(* IEC 61131-3 sources: canworks/library/modbus, 29 files *)

(* ---- CW_CHAR.st ---- *)
FUNCTION CW_CHAR : STRING
(* The one-character STRING of byte CODE ('' for 0), for building a STRING
   from bytes in plain ST: a look-up in tables of every byte value, 32 per
   table so that each fits the shortest default STRING length. *)
VAR_INPUT
  CODE : BYTE;
END_VAR
VAR
  t0 : STRING := '$01$02$03$04$05$06$07$08$09$0A$0B$0C$0D$0E$0F$10$11$12$13$14$15$16$17$18$19$1A$1B$1C$1D$1E$1F';
  t1 : STRING := '$20$21$22$23$24$25$26$27$28$29$2A$2B$2C$2D$2E$2F$30$31$32$33$34$35$36$37$38$39$3A$3B$3C$3D$3E$3F';
  t2 : STRING := '$40$41$42$43$44$45$46$47$48$49$4A$4B$4C$4D$4E$4F$50$51$52$53$54$55$56$57$58$59$5A$5B$5C$5D$5E$5F';
  t3 : STRING := '$60$61$62$63$64$65$66$67$68$69$6A$6B$6C$6D$6E$6F$70$71$72$73$74$75$76$77$78$79$7A$7B$7C$7D$7E$7F';
  t4 : STRING := '$80$81$82$83$84$85$86$87$88$89$8A$8B$8C$8D$8E$8F$90$91$92$93$94$95$96$97$98$99$9A$9B$9C$9D$9E$9F';
  t5 : STRING := '$A0$A1$A2$A3$A4$A5$A6$A7$A8$A9$AA$AB$AC$AD$AE$AF$B0$B1$B2$B3$B4$B5$B6$B7$B8$B9$BA$BB$BC$BD$BE$BF';
  t6 : STRING := '$C0$C1$C2$C3$C4$C5$C6$C7$C8$C9$CA$CB$CC$CD$CE$CF$D0$D1$D2$D3$D4$D5$D6$D7$D8$D9$DA$DB$DC$DD$DE$DF';
  t7 : STRING := '$E0$E1$E2$E3$E4$E5$E6$E7$E8$E9$EA$EB$EC$ED$EE$EF$F0$F1$F2$F3$F4$F5$F6$F7$F8$F9$FA$FB$FC$FD$FE$FF';
  k : INT;
END_VAR
k := BYTE_TO_INT(CODE);
CASE k / 32 OF
  0:
    IF k > 0 THEN
      CW_CHAR := MID(t0, 1, k);
    ELSE
      CW_CHAR := '';
    END_IF;
  1: CW_CHAR := MID(t1, 1, k MOD 32 + 1);
  2: CW_CHAR := MID(t2, 1, k MOD 32 + 1);
  3: CW_CHAR := MID(t3, 1, k MOD 32 + 1);
  4: CW_CHAR := MID(t4, 1, k MOD 32 + 1);
  5: CW_CHAR := MID(t5, 1, k MOD 32 + 1);
  6: CW_CHAR := MID(t6, 1, k MOD 32 + 1);
ELSE
  CW_CHAR := MID(t7, 1, k MOD 32 + 1);
END_CASE;
END_FUNCTION

FUNCTION CW_CHAR_CODE : BYTE
(* The byte value of the first character of C (0 for ''). *)
VAR_INPUT
  C : STRING;
END_VAR
VAR
  t0 : STRING := '$01$02$03$04$05$06$07$08$09$0A$0B$0C$0D$0E$0F$10$11$12$13$14$15$16$17$18$19$1A$1B$1C$1D$1E$1F';
  t1 : STRING := '$20$21$22$23$24$25$26$27$28$29$2A$2B$2C$2D$2E$2F$30$31$32$33$34$35$36$37$38$39$3A$3B$3C$3D$3E$3F';
  t2 : STRING := '$40$41$42$43$44$45$46$47$48$49$4A$4B$4C$4D$4E$4F$50$51$52$53$54$55$56$57$58$59$5A$5B$5C$5D$5E$5F';
  t3 : STRING := '$60$61$62$63$64$65$66$67$68$69$6A$6B$6C$6D$6E$6F$70$71$72$73$74$75$76$77$78$79$7A$7B$7C$7D$7E$7F';
  t4 : STRING := '$80$81$82$83$84$85$86$87$88$89$8A$8B$8C$8D$8E$8F$90$91$92$93$94$95$96$97$98$99$9A$9B$9C$9D$9E$9F';
  t5 : STRING := '$A0$A1$A2$A3$A4$A5$A6$A7$A8$A9$AA$AB$AC$AD$AE$AF$B0$B1$B2$B3$B4$B5$B6$B7$B8$B9$BA$BB$BC$BD$BE$BF';
  t6 : STRING := '$C0$C1$C2$C3$C4$C5$C6$C7$C8$C9$CA$CB$CC$CD$CE$CF$D0$D1$D2$D3$D4$D5$D6$D7$D8$D9$DA$DB$DC$DD$DE$DF';
  t7 : STRING := '$E0$E1$E2$E3$E4$E5$E6$E7$E8$E9$EA$EB$EC$ED$EE$EF$F0$F1$F2$F3$F4$F5$F6$F7$F8$F9$FA$FB$FC$FD$FE$FF';
  first : STRING;
  p : INT;
END_VAR
CW_CHAR_CODE := BYTE#0;
IF LEN(C) = 0 THEN
  RETURN;
END_IF;
first := LEFT(C, 1);
p := FIND(t0, first);
IF p > 0 THEN
  CW_CHAR_CODE := INT_TO_BYTE(p);
  RETURN;
END_IF;
p := FIND(t1, first);
IF p > 0 THEN
  CW_CHAR_CODE := INT_TO_BYTE(31 + p);
  RETURN;
END_IF;
p := FIND(t2, first);
IF p > 0 THEN
  CW_CHAR_CODE := INT_TO_BYTE(63 + p);
  RETURN;
END_IF;
p := FIND(t3, first);
IF p > 0 THEN
  CW_CHAR_CODE := INT_TO_BYTE(95 + p);
  RETURN;
END_IF;
p := FIND(t4, first);
IF p > 0 THEN
  CW_CHAR_CODE := INT_TO_BYTE(127 + p);
  RETURN;
END_IF;
p := FIND(t5, first);
IF p > 0 THEN
  CW_CHAR_CODE := INT_TO_BYTE(159 + p);
  RETURN;
END_IF;
p := FIND(t6, first);
IF p > 0 THEN
  CW_CHAR_CODE := INT_TO_BYTE(191 + p);
  RETURN;
END_IF;
p := FIND(t7, first);
IF p > 0 THEN
  CW_CHAR_CODE := INT_TO_BYTE(223 + p);
END_IF;
END_FUNCTION

(* ---- CW_REAL.st ---- *)
FUNCTION CW_DWORD_TO_REAL : REAL
(* The REAL whose IEEE 754 bit pattern is IN (a 32-bit value read from two
   Modbus registers). Infinities come back as +/-3.4E38, NaN as 0.0. *)
VAR_INPUT
  IN : DWORD;
END_VAR
VAR
  e : INT;
  m : LREAL;
  x : LREAL;
END_VAR
e := DWORD_TO_INT(SHR(IN, 23) AND DWORD#16#FF);
m := UDINT_TO_LREAL(DWORD_TO_UDINT(IN AND DWORD#16#7FFFFF));
IF e = 255 THEN
  IF m <> 0.0 THEN
    x := 0.0;
  ELSE
    x := 3.4028234663852886E38;
  END_IF;
ELSIF e = 0 THEN
  x := m * EXPT(2.0, -149);
ELSE
  x := (m + 8388608.0) * EXPT(2.0, e - 150);
END_IF;
IF (IN AND DWORD#16#80000000) <> DWORD#0 THEN
  x := -x;
END_IF;
CW_DWORD_TO_REAL := LREAL_TO_REAL(x);
END_FUNCTION

FUNCTION CW_REAL_TO_DWORD : DWORD
(* The IEEE 754 bit pattern of IN, to send a REAL in two Modbus registers. *)
VAR_INPUT
  IN : REAL;
END_VAR
VAR
  a : LREAL;
  e : INT;
  sign : DWORD;
END_VAR
a := REAL_TO_LREAL(IN);
sign := DWORD#0;
IF a < 0.0 THEN
  sign := DWORD#16#80000000;
  a := -a;
END_IF;
IF a <> a THEN
  CW_REAL_TO_DWORD := DWORD#16#7FC00000;
  RETURN;
END_IF;
IF a = 0.0 THEN
  CW_REAL_TO_DWORD := sign;
  RETURN;
END_IF;
IF a > 3.4028234663852886E38 THEN
  CW_REAL_TO_DWORD := sign OR DWORD#16#7F800000;
  RETURN;
END_IF;
e := LREAL_TO_INT(TRUNC(LN(a) / LN(2.0)));
WHILE a / EXPT(2.0, e) >= 2.0 DO
  e := e + 1;
END_WHILE;
WHILE a / EXPT(2.0, e) < 1.0 DO
  e := e - 1;
END_WHILE;
IF e < -126 THEN
  CW_REAL_TO_DWORD := sign OR UDINT_TO_DWORD(LREAL_TO_UDINT(a * EXPT(2.0, 149)));
ELSE
  CW_REAL_TO_DWORD := sign OR SHL(INT_TO_DWORD(e + 127), 23) OR UDINT_TO_DWORD(LREAL_TO_UDINT((a / EXPT(2.0, e) - 1.0) * 8388608.0));
END_IF;
END_FUNCTION

FUNCTION CW_LWORD_TO_LREAL : LREAL
(* The LREAL whose IEEE 754 bit pattern is IN (a 64-bit value read from four
   Modbus registers). Infinities come back as +/-1.79E308, NaN as 0.0. *)
VAR_INPUT
  IN : LWORD;
END_VAR
VAR
  e : INT;
  m : LREAL;
  x : LREAL;
END_VAR
e := LWORD_TO_INT(SHR(IN, 52) AND LWORD#16#7FF);
m := ULINT_TO_LREAL(LWORD_TO_ULINT(IN AND LWORD#16#FFFFFFFFFFFFF));
IF e = 2047 THEN
  IF m <> 0.0 THEN
    x := 0.0;
  ELSE
    x := 1.7976931348623157E308;
  END_IF;
ELSIF e = 0 THEN
  x := m * EXPT(2.0, -1074);
ELSE
  x := (m + 4503599627370496.0) * EXPT(2.0, e - 1075);
END_IF;
IF (IN AND SHL(LWORD#1, 63)) <> LWORD#0 THEN
  x := -x;
END_IF;
CW_LWORD_TO_LREAL := x;
END_FUNCTION

FUNCTION CW_LREAL_TO_LWORD : LWORD
(* The IEEE 754 bit pattern of IN, to send an LREAL in four Modbus registers. *)
VAR_INPUT
  IN : LREAL;
END_VAR
VAR
  a : LREAL;
  e : INT;
  sign : LWORD;
END_VAR
a := IN;
sign := LWORD#0;
IF a < 0.0 THEN
  sign := SHL(LWORD#1, 63);
  a := -a;
END_IF;
IF a <> a THEN
  CW_LREAL_TO_LWORD := LWORD#16#7FF8000000000000;
  RETURN;
END_IF;
IF a = 0.0 THEN
  CW_LREAL_TO_LWORD := sign;
  RETURN;
END_IF;
IF a > 1.7976931348623157E308 THEN
  CW_LREAL_TO_LWORD := sign OR LWORD#16#7FF0000000000000;
  RETURN;
END_IF;
e := LREAL_TO_INT(TRUNC(LN(a) / LN(2.0)));
WHILE a / EXPT(2.0, e) >= 2.0 DO
  e := e + 1;
END_WHILE;
WHILE a / EXPT(2.0, e) < 1.0 DO
  e := e - 1;
END_WHILE;
IF e < -1022 THEN
  CW_LREAL_TO_LWORD := sign OR ULINT_TO_LWORD(LREAL_TO_ULINT(a * EXPT(2.0, 537) * EXPT(2.0, 537)));
ELSE
  CW_LREAL_TO_LWORD := sign OR SHL(INT_TO_LWORD(e + 1023), 52) OR ULINT_TO_LWORD(LREAL_TO_ULINT((a / EXPT(2.0, e) - 1.0) * 4503599627370496.0));
END_IF;
END_FUNCTION

(* ---- CAN_BUS_INFO.st ---- *)
(*
 * CAN_BUS_INFO: the state of network NETWORK (one of the first 8) from the
 * bridge's network info block, updated every 100 ms, without a request:
 * STATE (0 error active, 1 warning, 2 error passive, 3 bus off, 4 unknown),
 * TX_ERRORS and RX_ERRORS (error counters), BUS_OFF_COUNT, BUS_LOAD (%),
 * RX_COUNT and TX_COUNT (frames), ERROR_FRAMES. ERROR_ID
 * (docs/plc-library.md#frame-blocks): 2 no such network, 20 the bridge is
 * not reachable, 22 the config has no network info (or NETWORK is past the
 * first 8).
 *)
(*
 * LINK is the generated `canworks.link` (ARRAY[0..1279] OF WORD); the block reads the bridge's network info block (see
 * CW_LINK_SERVICE for the words).
 *)
FUNCTION_BLOCK CAN_BUS_INFO
VAR_INPUT
  NETWORK : USINT;
END_VAR
VAR_IN_OUT
  LINK : ARRAY[0..1279] OF WORD;
END_VAR
VAR_OUTPUT
  STATE : USINT;
  TX_ERRORS : UINT;
  RX_ERRORS : UINT;
  BUS_OFF_COUNT : UDINT;
  BUS_LOAD : USINT;
  RX_COUNT : UDINT;
  TX_COUNT : UDINT;
  ERROR_FRAMES : UDINT;
  ERROR : BOOL;
  ERROR_ID : UINT;
END_VAR
VAR
  p : INT;
END_VAR
  ERROR_ID := 0;
  IF (LINK[21] AND WORD#16#0001) = WORD#0 THEN
    ERROR_ID := 20;
  ELSIF (LINK[89] AND WORD#16#0020) = WORD#0 OR NETWORK > 7 THEN
    ERROR_ID := 22;
  ELSE
    p := 960 + 18 * USINT_TO_INT(NETWORK);
    IF LINK[p + 17] = WORD#0 THEN
      ERROR_ID := 2;
    END_IF;
  END_IF;
  ERROR := ERROR_ID <> 0;
  IF ERROR THEN
    STATE := 4;
    TX_ERRORS := 0;
    RX_ERRORS := 0;
    BUS_OFF_COUNT := 0;
    BUS_LOAD := 0;
    RX_COUNT := 0;
    TX_COUNT := 0;
    ERROR_FRAMES := 0;
    RETURN;
  END_IF;
  STATE := WORD_TO_USINT(SHR(LINK[p], 8));
  BUS_LOAD := WORD_TO_USINT(LINK[p] AND WORD#16#00FF);
  TX_ERRORS := WORD_TO_UINT(LINK[p + 1]);
  RX_ERRORS := WORD_TO_UINT(LINK[p + 2]);
  BUS_OFF_COUNT := WORD_TO_UDINT(LINK[p + 3]) * 65536 + WORD_TO_UDINT(LINK[p + 4]);
  RX_COUNT := WORD_TO_UDINT(LINK[p + 5]) * 65536 + WORD_TO_UDINT(LINK[p + 6]);
  TX_COUNT := WORD_TO_UDINT(LINK[p + 7]) * 65536 + WORD_TO_UDINT(LINK[p + 8]);
  ERROR_FRAMES := WORD_TO_UDINT(LINK[p + 9]) * 65536 + WORD_TO_UDINT(LINK[p + 10]);
END_FUNCTION_BLOCK

(* ---- CAN_RECEIVE.st ---- *)
(*
 * CAN_RECEIVE: receives the CAN frames of network NETWORK whose identifier
 * matches ID under MASK (MASK 0: ID exactly; ALL_IDS: every frame of that
 * format), standard or EXTENDED, through a receiver of the bridge with a
 * queue of DEPTH frames (0: 32, at most 256). ENABLE opens it. Each call
 * gives at most one frame, oldest first: RECEIVED with RX_ID, RX_EXTENDED,
 * RX_RTR, RX_DLC, RX_DATA and TIMESTAMP (UTC microseconds, the receive time
 * of the bridge's batch, which its frames share: about one poll); call it
 * again in the same scan to read more
 * (`WHILE rx.RECEIVED DO ... rx(...); END_WHILE`).
 * QUEUED frames still wait in the bridge, OVERFLOW the queue was full,
 * DROPPED frames lost. ERROR_ID (docs/plc-library.md#frame-blocks): 1 the
 * network is not running, 2 no such network, 3 invalid input, 5 no free
 * receiver, 8 the bridge closed the receiver (it opens again), 20 the
 * bridge is not reachable, 22 the config has no receive or request mailbox.
 * After 1, 8 and 20 it opens again by itself.
 *)
(*
 * LINK is the generated `canworks.link` (ARRAY[0..1279] OF WORD); the block uses the bridge's receive mailbox and, to open and close its receiver, a
 * request mailbox (see
 * CW_LINK_SERVICE for the words).
 *)
FUNCTION_BLOCK CAN_RECEIVE
VAR_INPUT
  ENABLE : BOOL;
  NETWORK : USINT;
  ID : UDINT;
  MASK : UDINT;
  ALL_IDS : BOOL;
  EXTENDED : BOOL;
  DEPTH : UINT;
END_VAR
VAR_IN_OUT
  RX_DATA : ARRAY[0..7] OF BYTE;
  LINK : ARRAY[0..1279] OF WORD;
END_VAR
VAR_OUTPUT
  ACTIVE : BOOL;
  RECEIVED : BOOL;
  RX_ID : UDINT;
  RX_EXTENDED : BOOL;
  RX_RTR : BOOL;
  RX_DLC : USINT;
  TIMESTAMP : ULINT;
  QUEUED : UINT;
  OVERFLOW : BOOL;
  DROPPED : UDINT;
  ERROR : BOOL;
  ERROR_ID : UINT;
END_VAR
VAR
  rx : CW_RX;
  prev : BOOL;
  was_active : BOOL;
  last_drop : WORD;
  id_mask : UDINT;
  rec : INT;
  i : INT;
END_VAR
  IF ENABLE AND NOT prev THEN
    QUEUED := 0;
    OVERFLOW := FALSE;
    DROPPED := 0;
  END_IF;
  prev := ENABLE;
  IF ALL_IDS THEN
    id_mask := 0;
  ELSIF MASK <> 0 THEN
    id_mask := MASK;
  ELSIF EXTENDED THEN
    id_mask := 16#1FFFFFFF;
  ELSE
    id_mask := 16#7FF;
  END_IF;
  rx(ENABLE := ENABLE, CHANGED := FALSE, NEXT := TRUE, KIND := 1, NETWORK := NETWORK,
     FLAGS := SEL(EXTENDED, USINT#0, USINT#1), DEPTH := DEPTH, ID := ID, MASK := id_mask, RETRY := DWORD#16#00100102,
     LINK := LINK);
  IF rx.ACTIVE AND NOT was_active THEN
    last_drop := WORD#0;
  END_IF;
  was_active := rx.ACTIVE;
  RECEIVED := rx.RECEIVED;
  IF RECEIVED THEN
    rec := rx.REC;
    QUEUED := WORD_TO_UINT(LINK[rec + 1]);
    DROPPED := DROPPED + WORD_TO_UDINT(DINT_TO_WORD(WORD_TO_DINT(LINK[rec + 2]) - WORD_TO_DINT(last_drop)));
    last_drop := LINK[rec + 2];
    OVERFLOW := (LINK[rec] AND WORD#16#0004) <> WORD#0;
    TIMESTAMP := LWORD_TO_ULINT(SHL(WORD_TO_LWORD(LINK[741]), 48) OR SHL(WORD_TO_LWORD(LINK[742]), 32) OR
                 SHL(WORD_TO_LWORD(LINK[743]), 16) OR WORD_TO_LWORD(LINK[744]));
    RX_ID := WORD_TO_UDINT(LINK[rec + 3]) * 65536 + WORD_TO_UDINT(LINK[rec + 4]);
    RX_EXTENDED := (LINK[rec + 5] AND WORD#16#0100) <> WORD#0;
    RX_RTR := (LINK[rec + 5] AND WORD#16#0200) <> WORD#0;
    RX_DLC := WORD_TO_USINT(LINK[rec + 5] AND WORD#16#00FF);
    FOR i := 0 TO 3 DO
      RX_DATA[2 * i] := WORD_TO_BYTE(SHR(LINK[rec + 6 + i], 8));
      RX_DATA[2 * i + 1] := WORD_TO_BYTE(LINK[rec + 6 + i]);
    END_FOR;
  END_IF;
  ACTIVE := rx.ACTIVE;
  ERROR := rx.ERROR;
  ERROR_ID := rx.ERROR_ID;
END_FUNCTION_BLOCK

(* ---- CAN_SEND.st ---- *)
(*
 * CAN_SEND: sends one CAN frame (ID, EXTENDED, RTR, DLC 0..8 bytes of DATA)
 * on network NETWORK. A rising edge of EXECUTE starts it; BUSY until the
 * bridge has sent it, then DONE or ERROR with ERROR_ID
 * (docs/plc-library.md#frame-blocks): 1 the network is not running, 2 no
 * such network, 3 invalid input, 5 too many frames wait, 6 not sent within
 * TIMEOUT (T#0s: 1 s), 7 the bus is off, 8 cancelled, 20 the bridge is not
 * reachable, 22 the config has no request mailbox.
 *)
(*
 * LINK is the generated `canworks.link` (ARRAY[0..1279] OF WORD); the block uses a request mailbox of the bridge (`mailboxes` in the config); instances share
 * them in the order they started (see
 * CW_LINK_SERVICE for the words).
 *)
FUNCTION_BLOCK CAN_SEND
VAR_INPUT
  EXECUTE : BOOL;
  NETWORK : USINT;
  ID : UDINT;
  EXTENDED : BOOL;
  RTR : BOOL;
  DLC : USINT;
  TIMEOUT : TIME;
END_VAR
VAR_IN_OUT
  DATA : ARRAY[0..7] OF BYTE;
  LINK : ARRAY[0..1279] OF WORD;
END_VAR
VAR_OUTPUT
  BUSY : BOOL;
  DONE : BOOL;
  ERROR : BOOL;
  ERROR_ID : UINT;
END_VAR
VAR
  x : CW_REQUEST;
  buf : ARRAY[0..1784] OF BYTE;
  prev : BOOL;
  refused : UINT;
  flags : WORD;
  ms : UDINT;
  i : INT;
END_VAR
  IF EXECUTE AND NOT prev AND NOT x.BUSY THEN
    refused := 0;
    IF DLC > 8 THEN
      refused := 3;
    END_IF;
    FOR i := 0 TO 7 DO
      buf[i] := DATA[i];
    END_FOR;
  ELSIF NOT EXECUTE THEN
    refused := 0;
  END_IF;
  prev := EXECUTE;
  flags := SEL(EXTENDED, WORD#0, WORD#1) OR SEL(RTR, WORD#0, WORD#2);
  ms := DWORD_TO_UDINT(TIME_TO_DWORD(TIMEOUT));
  IF ms > 65535 THEN
    ms := 65535;
  END_IF;
  x(EXECUTE := EXECUTE AND refused = 0, OP := 5, NET := NETWORK, A0 := DWORD_TO_WORD(SHR(UDINT_TO_DWORD(ID), 16)),
    A1 := UDINT_TO_WORD(ID), A2 := SHL(flags, 8) OR USINT_TO_WORD(DLC), A3 := UDINT_TO_WORD(ms), A4 := WORD#0, A5 := WORD#0,
    LENGTH := 8, FETCH_MAX := 0, LINK := LINK, DATA := buf);
  BUSY := x.BUSY;
  DONE := x.DONE;
  ERROR := x.ERROR OR refused <> 0;
  ERROR_ID := SEL(refused <> 0, x.ERROR_ID, refused);
END_FUNCTION_BLOCK

(* ---- CAN_SEND_CYCLIC.st ---- *)
(*
 * CAN_SEND_CYCLIC: the bridge sends one CAN frame (ID, EXTENDED, DLC bytes
 * of DATA) on network NETWORK every PERIOD (1 ms .. 60 s) while ENABLE is
 * TRUE. Changed DATA, DLC or PERIOD go to the bridge when they change; the
 * block must be called at least every second (its keepalive), or the bridge
 * stops the frame. ACTIVE while the job runs, COUNT frames sent. ERROR_ID
 * (docs/plc-library.md#frame-blocks): 1 the network is not running, 2 no
 * such network, 3 invalid input, 5 no free cyclic job, 7 the bus is off
 * (the job stays), 8 cancelled (the bridge stopped the job; it starts
 * again), 20 the bridge is not reachable, 22 the config has no request
 * mailbox or no cyclic jobs. After 1, 7, 8 and 20 it starts again by itself.
 *)
(*
 * LINK is the generated `canworks.link` (ARRAY[0..1279] OF WORD); the block uses a request mailbox of the bridge (`mailboxes` in the config); instances share
 * them in the order they started, and a cyclic job of the bridge's table (see
 * CW_LINK_SERVICE for the words).
 *)
FUNCTION_BLOCK CAN_SEND_CYCLIC
VAR_INPUT
  ENABLE : BOOL;
  NETWORK : USINT;
  ID : UDINT;
  EXTENDED : BOOL;
  DLC : USINT;
  PERIOD : TIME;
END_VAR
VAR_IN_OUT
  DATA : ARRAY[0..7] OF BYTE;
  LINK : ARRAY[0..1279] OF WORD;
END_VAR
VAR_OUTPUT
  ACTIVE : BOOL;
  COUNT : UDINT;
  ERROR : BOOL;
  ERROR_ID : UINT;
END_VAR
VAR
  mb : CW_MB_CALL;
  prev : BOOL;
  phase : USINT;           (* 0 off, 1 starting, 2 running, 3 updating, 4 stopping *)
  job : INT;
  gen : WORD;
  tick0 : WORD;
  sent : ARRAY[0..7] OF BYTE;
  sent_dlc : USINT;
  sent_ms : UDINT;
  ms : UDINT;
  changed : BOOL;
  t : INT;
  i : INT;
  err : UINT;
  fresh : BOOL;
END_VAR
  err := 0;
  ms := DWORD_TO_UDINT(TIME_TO_DWORD(PERIOD));
  IF ms > 65535 THEN
    ms := 65535;
  END_IF;
  IF ENABLE AND NOT prev THEN
    COUNT := 0;
    ERROR := FALSE;
    ERROR_ID := 0;
  END_IF;
  IF (LINK[21] AND WORD#16#0001) = WORD#0 AND phase <> 0 THEN
    mb(RUN := FALSE, LINK := LINK);
    phase := 0;
    IF ENABLE THEN
      err := 20;
    END_IF;
  END_IF;
  IF phase = 2 OR phase = 3 THEN
    LINK[128 + job] := UDINT_TO_WORD(WORD_TO_UDINT(LINK[128 + job]) + 1);
    t := 1105 + 4 * job;
    fresh := (DINT_TO_WORD(WORD_TO_DINT(LINK[1104]) - WORD_TO_DINT(tick0)) AND WORD#16#8000) = WORD#0;
    IF fresh AND LINK[t + 1] <> gen THEN
      mb(RUN := FALSE, LINK := LINK);
      phase := 0;
      err := 8;
    ELSIF fresh THEN
      COUNT := WORD_TO_UDINT(LINK[t + 2]) * 65536 + WORD_TO_UDINT(LINK[t + 3]);
      IF SHR(LINK[t], 8) = WORD#2 THEN
        ERROR := TRUE;
        ERROR_ID := WORD_TO_UINT(LINK[t] AND WORD#16#00FF);
      ELSIF ERROR AND ERROR_ID = 7 THEN
        ERROR := FALSE;
        ERROR_ID := 0;
      END_IF;
    END_IF;
  END_IF;
  IF (phase = 2 OR phase = 3) AND NOT ENABLE THEN
    phase := 4;
  END_IF;
  changed := DLC <> sent_dlc OR ms <> sent_ms;
  FOR i := 0 TO 7 DO
    IF DATA[i] <> sent[i] THEN
      changed := TRUE;
    END_IF;
  END_FOR;
  IF phase = 2 AND changed THEN
    phase := 3;
  END_IF;
  IF phase = 0 AND ENABLE AND err = 0 AND
     NOT (ERROR AND ERROR_ID <> 1 AND ERROR_ID <> 7 AND ERROR_ID <> 8 AND ERROR_ID <> 20) THEN
    ERROR := FALSE;
    ERROR_ID := 0;
    IF (LINK[21] AND WORD#16#0001) = WORD#0 THEN
      err := 20;
    ELSIF (LINK[89] AND WORD#16#0007) = WORD#0 OR (LINK[89] AND WORD#16#1F00) = WORD#0 THEN
      err := 22;
    ELSIF DLC > 8 THEN
      err := 3;
    ELSE
      phase := 1;
    END_IF;
  END_IF;
  IF phase = 1 OR phase = 3 OR phase = 4 THEN
    mb(RUN := TRUE, SEND := FALSE, LINK := LINK);
    IF mb.LOST THEN
      phase := 0;
      err := SEL(ENABLE, UINT#0, UINT#20);
    ELSIF mb.ANSWERED THEN
      IF phase = 4 THEN
        phase := 0;
      ELSIF mb.ERR <> 0 THEN
        err := mb.ERR;
        IF phase = 1 OR mb.ERR = 8 THEN
          phase := 0;
        ELSE
          phase := 2;
        END_IF;
      ELSE
        IF phase = 1 THEN
          job := WORD_TO_INT(LINK[mb.BASE + 74]);
          gen := LINK[mb.BASE + 75];
          tick0 := LINK[mb.BASE + 76];
          COUNT := 0;
        END_IF;
        phase := 2;
      END_IF;
      mb(RUN := FALSE, LINK := LINK);
    ELSIF mb.OWNED AND NOT mb.WAITING THEN
      IF phase = 4 THEN
        mb(RUN := TRUE, SEND := TRUE, OP := 7, NET := NETWORK, A0 := INT_TO_WORD(job), A1 := WORD#0, A2 := WORD#0, A3 := WORD#0,
           A4 := WORD#0, A5 := WORD#0, LINK := LINK);
      ELSE
        FOR i := 0 TO 3 DO
          LINK[mb.BASE + 8 + i] := SHL(BYTE_TO_WORD(DATA[2 * i]), 8) OR BYTE_TO_WORD(DATA[2 * i + 1]);
          sent[2 * i] := DATA[2 * i];
          sent[2 * i + 1] := DATA[2 * i + 1];
        END_FOR;
        sent_dlc := DLC;
        sent_ms := ms;
        mb(RUN := TRUE, SEND := TRUE, OP := 6, NET := NETWORK, A0 := SEL(phase = 1, INT_TO_WORD(job), WORD#16#FFFF),
           A1 := DWORD_TO_WORD(SHR(UDINT_TO_DWORD(ID), 16)), A2 := UDINT_TO_WORD(ID),
           A3 := SHL(SEL(EXTENDED, WORD#0, WORD#1), 8) OR USINT_TO_WORD(DLC), A4 := UDINT_TO_WORD(ms), A5 := WORD#0,
           LINK := LINK);
      END_IF;
    END_IF;
  END_IF;
  IF err <> 0 THEN
    ERROR := TRUE;
    ERROR_ID := err;
  END_IF;
  ACTIVE := phase = 2 OR phase = 3;
  prev := ENABLE;
END_FUNCTION_BLOCK

(* ---- CO_NMT.st ---- *)
(*
 * CO_NMT: sends the NMT command COMMAND (CiA 301 codes: 1 START, 2 STOP,
 * 128 ENTER PRE-OPERATIONAL, 129 RESET NODE, 130 RESET COMMUNICATION) to
 * node NODE (0: every node) of CANopen master network NETWORK, through the
 * bridge's control block. A rising edge of EXECUTE starts it; BUSY until the
 * bridge has handled it, then DONE or ERROR with ERROR_ID (docs/plc-library.md):
 * 2 no answer within TIMEOUT (T#0s: 5 s), 5 refused (the bus is down or 16
 * commands wait), 6 invalid input, 20 the bridge is not reachable, 22 the
 * config has no control block, 8 cancelled: the bridge restarted and did
 * not run it (start it again). Instances share the control block: one waits
 * while another uses it.
 *)
(*
 * LINK is the generated `canworks.link` (ARRAY[0..1279] OF WORD): the
 * bridge's blocks as canworks_in and canworks_out copy them from and to the
 * Modbus registers every scan, one word per register (high byte = the
 * bridge's even byte). Words: 0-3 status block, 4-6 control block, 7-13 SDO
 * request, 14-20 SDO response, 21 flags (bit 0 the bridge answers with this
 * program's map, 1 a control block, 2 SDO registers, 8 + n a live list for
 * network n), 22 control block owner, 23 SDO owner, 24 last instance number,
 * 25 + 8n .. 32 + 8n the live list of network n (n 0..7).
 *)
FUNCTION_BLOCK CO_NMT
VAR_INPUT
  EXECUTE : BOOL;
  NETWORK : USINT;
  NODE : USINT;
  COMMAND : USINT;
  TIMEOUT : TIME;
END_VAR
VAR_OUTPUT
  BUSY : BOOL;
  DONE : BOOL;
  ERROR : BOOL;
  ERROR_ID : UINT;
END_VAR
VAR_IN_OUT
  LINK : ARRAY[0..1279] OF WORD;
END_VAR
VAR
  me : WORD;
  prev : BOOL;
  phase : USINT;           (* 0 idle, 1 waiting for the control block, 2 sent, 3 ended *)
  cmd : WORD;
  counter : WORD;
  timer : TON;
  result : WORD;
  err : UINT;
  fin : BOOL;
END_VAR
  IF me = WORD#0 THEN
    LINK[24] := UINT_TO_WORD(WORD_TO_UINT(LINK[24]) + 1);
    me := LINK[24];
  END_IF;
  IF phase = 3 AND NOT EXECUTE THEN
    phase := 0;
    DONE := FALSE;
    ERROR := FALSE;
  END_IF;
  err := 0;
  fin := FALSE;
  IF phase = 0 AND EXECUTE AND NOT prev THEN
    DONE := FALSE;
    ERROR := FALSE;
    ERROR_ID := 0;
    timer(IN := FALSE);
    CASE COMMAND OF
      1: cmd := WORD#3;
      2: cmd := WORD#4;
      128: cmd := WORD#5;
      129: cmd := WORD#6;
      130: cmd := WORD#7;
    ELSE
      cmd := WORD#0;
    END_CASE;
    IF (LINK[21] AND WORD#16#0001) = WORD#0 THEN
      err := 20;
    ELSIF (LINK[21] AND WORD#16#0002) = WORD#0 THEN
      err := 22;
    ELSIF cmd = WORD#0 OR NODE > 127 THEN
      err := 6;
    ELSE
      phase := 1;
    END_IF;
  END_IF;
  IF phase = 1 OR phase = 2 THEN
    timer(IN := TRUE, PT := SEL(TIMEOUT = T#0s, TIMEOUT, T#5s));
    IF (LINK[21] AND WORD#16#0001) = WORD#0 THEN
      err := 20;
    ELSIF timer.Q THEN
      err := 2;
    ELSIF phase = 1 AND (LINK[22] = WORD#0 OR LINK[22] = me) THEN
      LINK[22] := me;
      counter := UINT_TO_WORD(WORD_TO_UINT(LINK[2]) + 1);
      LINK[4] := counter;
      LINK[5] := SHL(cmd, 8) OR USINT_TO_WORD(NETWORK);
      LINK[6] := SHL(USINT_TO_WORD(NODE), 8);
      phase := 2;
    ELSIF phase = 2 AND LINK[2] = counter THEN
      result := SHR(LINK[3], 8);
      IF result = WORD#0 THEN
        fin := TRUE;
      ELSIF result = WORD#5 THEN
        err := 5;
      ELSIF result = WORD#6 THEN
        err := 8;              (* the bridge restarted and did not run it *)
      ELSE
        err := 6;
      END_IF;
    END_IF;
  END_IF;
  IF err <> 0 OR fin THEN
    phase := 3;
    DONE := fin;
    ERROR := err <> 0;
    ERROR_ID := err;
    timer(IN := FALSE);
    IF LINK[22] = me THEN
      LINK[22] := WORD#0;
    END_IF;
  END_IF;
  BUSY := phase = 1 OR phase = 2;
  prev := EXECUTE;
END_FUNCTION_BLOCK

(* ---- CO_NODE_LIVE.st ---- *)
(*
 * CO_NODE_LIVE: TRUE while node NODE of CANopen master network NETWORK is
 * OPERATIONAL, from the bridge's live list of that network. FALSE without a
 * live list for the network or while the bridge is not reachable.
 *)
(*
 * LINK is the generated `canworks.link` (ARRAY[0..1279] OF WORD): the
 * bridge's blocks as canworks_in and canworks_out copy them from and to the
 * Modbus registers every scan, one word per register (high byte = the
 * bridge's even byte). Words: 0-3 status block, 4-6 control block, 7-13 SDO
 * request, 14-20 SDO response, 21 flags (bit 0 the bridge answers with this
 * program's map, 1 a control block, 2 SDO registers, 8 + n a live list for
 * network n), 22 control block owner, 23 SDO owner, 24 last instance number,
 * 25 + 8n .. 32 + 8n the live list of network n (n 0..7).
 *)
FUNCTION_BLOCK CO_NODE_LIVE
VAR_INPUT
  NETWORK : USINT;
  NODE : USINT;
END_VAR
VAR_OUTPUT
  LIVE : BOOL;
END_VAR
VAR_IN_OUT
  LINK : ARRAY[0..1279] OF WORD;
END_VAR
VAR
  byte_no : INT;
  wd : WORD;
  bit_no : INT;
END_VAR
  LIVE := FALSE;
  IF (LINK[21] AND WORD#16#0001) <> WORD#0 AND NETWORK < 8 AND NODE >= 1 AND NODE <= 127 THEN
    IF (SHR(LINK[21], USINT_TO_UINT(NETWORK) + 8) AND WORD#16#0001) <> WORD#0 THEN
      byte_no := USINT_TO_INT(NODE) / 8;
      wd := LINK[25 + USINT_TO_INT(NETWORK) * 8 + byte_no / 2];
      bit_no := USINT_TO_INT(NODE) MOD 8;
      IF byte_no MOD 2 = 0 THEN
        bit_no := bit_no + 8;
      END_IF;
      LIVE := (SHR(wd, INT_TO_UINT(bit_no)) AND WORD#16#0001) <> WORD#0;
    END_IF;
  END_IF;
END_FUNCTION_BLOCK

(* ---- CO_RECV_EMCY.st ---- *)
(*
 * CO_RECV_EMCY: receives the EMCY messages of node NODE (0: every node) of
 * CANopen master network NETWORK from the bridge's EMCY history, from the
 * oldest kept message or, with SKIP_OLD, from the next one. ENABLE starts
 * it. Each call gives at most one message, oldest first: RECEIVED with
 * EMCY_NODE, ERROR_CODE, ERROR_REGISTER, MSEF (5 manufacturer bytes) and
 * TIMESTAMP (UTC microseconds). QUEUED messages still wait, LOST messages
 * the history dropped before they were read (OVERFLOW then TRUE).
 * ERROR_ID (docs/plc-library.md#sdo-blocks): 4 the network is not running
 * (tried again), 5 no free receiver, 6 invalid input, 8 a new CANopen
 * session (shown for one call, reading goes on with the new session's
 * messages) or the bridge closed the receiver (it starts again), 20 the
 * bridge is not reachable, 22 the config has no receive or request mailbox.
 *)
(*
 * LINK is the generated `canworks.link` (ARRAY[0..1279] OF WORD); the block uses the bridge's receive mailbox and a request mailbox (see
 * CW_LINK_SERVICE for the words).
 *)
FUNCTION_BLOCK CO_RECV_EMCY
VAR_INPUT
  ENABLE : BOOL;
  NETWORK : USINT;
  NODE : USINT;
  SKIP_OLD : BOOL;
END_VAR
VAR_IN_OUT
  MSEF : ARRAY[0..4] OF BYTE;
  LINK : ARRAY[0..1279] OF WORD;
END_VAR
VAR_OUTPUT
  ACTIVE : BOOL;
  RECEIVED : BOOL;
  EMCY_NODE : USINT;
  ERROR_CODE : WORD;
  ERROR_REGISTER : BYTE;
  TIMESTAMP : ULINT;
  QUEUED : UINT;
  OVERFLOW : BOOL;
  LOST : UDINT;
  ERROR : BOOL;
  ERROR_ID : UINT;
END_VAR
VAR
  rx : CW_RX;
  prev : BOOL;
  was_active : BOOL;
  last_drop : WORD;
  lost_now : UDINT;
  restart : BOOL;
  rec : INT;
END_VAR
  RECEIVED := FALSE;
  restart := FALSE;
  IF ENABLE AND NOT prev THEN
    QUEUED := 0;
    OVERFLOW := FALSE;
    LOST := 0;
  ELSIF NOT ENABLE AND prev THEN
    QUEUED := 0;
    OVERFLOW := FALSE;
  END_IF;
  prev := ENABLE;
  rx(ENABLE := ENABLE, CHANGED := FALSE, NEXT := TRUE, KIND := 3, NETWORK := NETWORK,
     FLAGS := SEL(SKIP_OLD, USINT#0, USINT#1), DEPTH := 0, ID := 0, MASK := USINT_TO_UDINT(NODE),
     RETRY := DWORD#16#00100110, LINK := LINK);
  IF rx.ACTIVE AND NOT was_active THEN
    last_drop := WORD#0;
  END_IF;
  was_active := rx.ACTIVE;
  IF rx.RECEIVED THEN
    rec := rx.REC;
    QUEUED := WORD_TO_UINT(LINK[rec + 1]);
    lost_now := WORD_TO_UDINT(DINT_TO_WORD(WORD_TO_DINT(LINK[rec + 2]) - WORD_TO_DINT(last_drop)));
    last_drop := LINK[rec + 2];
    LOST := LOST + lost_now;
    IF lost_now <> 0 THEN
      OVERFLOW := TRUE;
    END_IF;
    IF (LINK[rec] AND WORD#16#0002) <> WORD#0 THEN
      restart := TRUE;
    ELSE
      RECEIVED := TRUE;
      TIMESTAMP := LWORD_TO_ULINT(SHL(WORD_TO_LWORD(LINK[rec + 3]), 48) OR SHL(WORD_TO_LWORD(LINK[rec + 4]), 32) OR
                   SHL(WORD_TO_LWORD(LINK[rec + 5]), 16) OR WORD_TO_LWORD(LINK[rec + 6]));
      EMCY_NODE := WORD_TO_USINT(SHR(LINK[rec + 7], 8));
      ERROR_REGISTER := WORD_TO_BYTE(LINK[rec + 7]);
      ERROR_CODE := LINK[rec + 8];
      MSEF[0] := WORD_TO_BYTE(SHR(LINK[rec + 9], 8));
      MSEF[1] := WORD_TO_BYTE(LINK[rec + 9]);
      MSEF[2] := WORD_TO_BYTE(SHR(LINK[rec + 10], 8));
      MSEF[3] := WORD_TO_BYTE(LINK[rec + 10]);
      MSEF[4] := WORD_TO_BYTE(SHR(LINK[rec + 11], 8));
    END_IF;
  END_IF;
  ACTIVE := rx.ACTIVE;
  ERROR := rx.ERROR OR restart;
  ERROR_ID := SEL(restart, rx.ERROR_ID, UINT#8);
END_FUNCTION_BLOCK

(* ---- CO_SDO_READ.st ---- *)
(*
 * CO_SDO_READ: reads object INDEX:SUBINDEX (up to 4 bytes) of node NODE
 * (1..127) of CANopen master network NETWORK into DATA, through the bridge's
 * SDO registers.
 * A rising edge of EXECUTE starts it; BUSY until the bridge has an answer,
 * then DONE or ERROR with ERROR_ID (docs/plc-library.md): 1 the node aborted
 * (ABORT_CODE), 2 no answer within TIMEOUT (T#0s: 5 s), 6 invalid input,
 * 20 the bridge is not reachable, 21 SDO writes are not allowed by the
 * config (ABORT_CODE 16#08000020), 22 the config has no SDO registers,
 * 8 cancelled: the bridge restarted and did not send it (start it again).
 * Instances share the SDO registers: one waits while another uses them.
 *)
(*
 * LINK is the generated `canworks.link` (ARRAY[0..1279] OF WORD): the
 * bridge's blocks as canworks_in and canworks_out copy them from and to the
 * Modbus registers every scan, one word per register (high byte = the
 * bridge's even byte). Words: 0-3 status block, 4-6 control block, 7-13 SDO
 * request, 14-20 SDO response, 21 flags (bit 0 the bridge answers with this
 * program's map, 1 a control block, 2 SDO registers, 8 + n a live list for
 * network n), 22 control block owner, 23 SDO owner, 24 last instance number,
 * 25 + 8n .. 32 + 8n the live list of network n (n 0..7).
 *)
FUNCTION_BLOCK CO_SDO_READ
VAR_INPUT
  EXECUTE : BOOL;
  NETWORK : USINT;
  NODE : USINT;
  INDEX : UINT;
  SUBINDEX : USINT;
  TIMEOUT : TIME;
END_VAR
VAR_OUTPUT
  BUSY : BOOL;
  DONE : BOOL;
  ERROR : BOOL;
  ERROR_ID : UINT;
  ABORT_CODE : UDINT;
  DATA : UDINT;
END_VAR
VAR_IN_OUT
  LINK : ARRAY[0..1279] OF WORD;
END_VAR
VAR
  me : WORD;
  prev : BOOL;
  phase : USINT;           (* 0 idle, 1 waiting for the SDO registers, 2 sent, 3 ended *)
  counter : WORD;
  timer : TON;
  state : WORD;
  err : UINT;
  fin : BOOL;
END_VAR
  IF me = WORD#0 THEN
    LINK[24] := UINT_TO_WORD(WORD_TO_UINT(LINK[24]) + 1);
    me := LINK[24];
  END_IF;
  IF phase = 3 AND NOT EXECUTE THEN
    phase := 0;
    DONE := FALSE;
    ERROR := FALSE;
  END_IF;
  err := 0;
  fin := FALSE;
  IF phase = 0 AND EXECUTE AND NOT prev THEN
    DONE := FALSE;
    ERROR := FALSE;
    ERROR_ID := 0;
    ABORT_CODE := 0;
    DATA := 0;
    timer(IN := FALSE);
    IF (LINK[21] AND WORD#16#0001) = WORD#0 THEN
      err := 20;
    ELSIF (LINK[21] AND WORD#16#0004) = WORD#0 THEN
      err := 22;
    ELSIF NODE < 1 OR NODE > 127 THEN
      err := 6;
    ELSE
      phase := 1;
    END_IF;
  END_IF;
  IF phase = 1 OR phase = 2 THEN
    timer(IN := TRUE, PT := SEL(TIMEOUT = T#0s, TIMEOUT, T#5s));
    IF (LINK[21] AND WORD#16#0001) = WORD#0 THEN
      err := 20;
    ELSIF timer.Q THEN
      err := 2;
      ABORT_CODE := 16#05040000;
    ELSIF phase = 1 AND (LINK[23] = WORD#0 OR LINK[23] = me) THEN
      LINK[23] := me;
      counter := UINT_TO_WORD(WORD_TO_UINT(LINK[14]) + 1);
      LINK[7] := counter;
      LINK[8] := SHL(WORD#1, 8) OR USINT_TO_WORD(NETWORK);
      LINK[9] := SHL(USINT_TO_WORD(NODE), 8) OR USINT_TO_WORD(SUBINDEX);
      LINK[10] := UINT_TO_WORD(INDEX);
      LINK[11] := WORD#0;
      LINK[12] := WORD#0;
      LINK[13] := WORD#0;
      phase := 2;
    ELSIF phase = 2 AND LINK[14] = counter THEN
      state := SHR(LINK[15], 8);
      IF state = WORD#2 THEN
        DATA := DWORD_TO_UDINT(SHL(WORD_TO_DWORD(LINK[18]), 16) OR WORD_TO_DWORD(LINK[19]));
        fin := TRUE;
      ELSIF state = WORD#3 THEN
        ABORT_CODE := DWORD_TO_UDINT(SHL(WORD_TO_DWORD(LINK[16]), 16) OR WORD_TO_DWORD(LINK[17]));
        IF ABORT_CODE = 16#08000020 THEN
          err := 21;
        ELSIF ABORT_CODE = 16#08000021 THEN
          err := 8;            (* the bridge restarted and did not send it *)
        ELSE
          err := 1;
        END_IF;
      END_IF;
    END_IF;
  END_IF;
  IF err <> 0 OR fin THEN
    phase := 3;
    DONE := fin;
    ERROR := err <> 0;
    ERROR_ID := err;
    timer(IN := FALSE);
    IF LINK[23] = me THEN
      LINK[23] := WORD#0;
    END_IF;
  END_IF;
  BUSY := phase = 1 OR phase = 2;
  prev := EXECUTE;
END_FUNCTION_BLOCK

(* ---- CO_SDO_READ_BYTES.st ---- *)
(*
 * CO_SDO_READ_BYTES: reads object INDEX:SUBINDEX of node NODE (1..127) of
 * CANopen master network NETWORK into BUFFER, up to 1024 bytes; SIZE is the
 * object's size.
 * A rising edge of EXECUTE starts it; BUSY until the bridge has an answer,
 * then DONE or ERROR with ERROR_ID (docs/plc-library.md#sdo-blocks): 1 the
 * node aborted (ABORT_CODE), 2 no answer within TIMEOUT (T#0s: 5 s), 4 the
 * network is not running, 5 too many SDO requests wait, 6 invalid input,
 * 7 too large (more than 1024 bytes; SIZE says how many), 8 cancelled, 20 the bridge is not reachable, 22 the config
 * has no request mailbox.
 *)
(*
 * LINK is the generated `canworks.link` (ARRAY[0..1279] OF WORD); the block
 * uses a request mailbox of the bridge (`mailboxes` in the config, see
 * CW_LINK_SERVICE for the words). Instances share the request mailboxes in
 * the order they started.
 *)
FUNCTION_BLOCK CO_SDO_READ_BYTES
VAR_INPUT
  EXECUTE : BOOL;
  NETWORK : USINT;
  NODE : USINT;
  INDEX : UINT;
  SUBINDEX : USINT;
  TIMEOUT : TIME;
END_VAR
VAR_OUTPUT
  BUSY : BOOL;
  DONE : BOOL;
  ERROR : BOOL;
  ERROR_ID : UINT;
  ABORT_CODE : UDINT;
  SIZE : UINT;
END_VAR
VAR_IN_OUT
  BUFFER : ARRAY[0..1023] OF BYTE;
  LINK : ARRAY[0..1279] OF WORD;
END_VAR
VAR
  x : CW_SDO_XFER;
END_VAR
  x(EXECUTE := EXECUTE, WRITE := FALSE, NETWORK := NETWORK, NODE := NODE, INDEX := INDEX, SUBINDEX := SUBINDEX,
    TIMEOUT := TIMEOUT, KIND := 3, MAX_SIZE := 1024, FETCH_MAX := 1024, LINK := LINK, DATA := BUFFER);
  BUSY := x.BUSY;
  DONE := x.DONE;
  ERROR := x.ERROR;
  ERROR_ID := x.ERROR_ID;
  ABORT_CODE := x.ABORT_CODE;
  IF x.RSIZE > 65535 THEN
    SIZE := 65535;
  ELSE
    SIZE := UDINT_TO_UINT(x.RSIZE);
  END_IF;
END_FUNCTION_BLOCK

(* ---- CO_SDO_READ_REAL.st ---- *)
(*
 * CO_SDO_READ_REAL: reads object INDEX:SUBINDEX (REAL32 or REAL64) of node
 * NODE (1..127) of CANopen master network NETWORK into VALUE.
 * A rising edge of EXECUTE starts it; BUSY until the bridge has an answer,
 * then DONE or ERROR with ERROR_ID (docs/plc-library.md#sdo-blocks): 1 the
 * node aborted (ABORT_CODE), 2 no answer within TIMEOUT (T#0s: 5 s), 4 the
 * network is not running, 5 too many SDO requests wait, 6 invalid input,
 * 7 too large (a reply that is not 4 or 8 bytes), 8 cancelled, 20 the bridge is not reachable, 22 the config
 * has no request mailbox.
 *)
(*
 * LINK is the generated `canworks.link` (ARRAY[0..1279] OF WORD); the block
 * uses a request mailbox of the bridge (`mailboxes` in the config, see
 * CW_LINK_SERVICE for the words). Instances share the request mailboxes in
 * the order they started.
 *)
FUNCTION_BLOCK CO_SDO_READ_REAL
VAR_INPUT
  EXECUTE : BOOL;
  NETWORK : USINT;
  NODE : USINT;
  INDEX : UINT;
  SUBINDEX : USINT;
  TIMEOUT : TIME;
END_VAR
VAR_OUTPUT
  BUSY : BOOL;
  DONE : BOOL;
  ERROR : BOOL;
  ERROR_ID : UINT;
  ABORT_CODE : UDINT;
  VALUE : LREAL;
END_VAR
VAR_IN_OUT
  LINK : ARRAY[0..1279] OF WORD;
END_VAR
VAR
  x : CW_SDO_XFER;
  buf : ARRAY[0..1023] OF BYTE;
  was : BOOL;
  bad : BOOL;
  bits : LWORD;
  i : INT;
END_VAR
  x(EXECUTE := EXECUTE, WRITE := FALSE, NETWORK := NETWORK, NODE := NODE, INDEX := INDEX, SUBINDEX := SUBINDEX,
    TIMEOUT := TIMEOUT, KIND := 1, MAX_SIZE := 8, FETCH_MAX := 8, LINK := LINK, DATA := buf);
  BUSY := x.BUSY;
  DONE := x.DONE;
  ERROR := x.ERROR;
  ERROR_ID := x.ERROR_ID;
  ABORT_CODE := x.ABORT_CODE;
  IF x.DONE AND NOT was THEN
    bad := x.RSIZE <> 4 AND x.RSIZE <> 8;
    IF NOT bad THEN
      bits := LWORD#0;
      FOR i := UDINT_TO_INT(x.RSIZE) - 1 TO 0 BY -1 DO
        bits := SHL(bits, 8) OR BYTE_TO_LWORD(buf[i]);
      END_FOR;
      IF x.RSIZE = 4 THEN
        VALUE := REAL_TO_LREAL(CW_DWORD_TO_REAL(LWORD_TO_DWORD(bits)));
      ELSE
        VALUE := CW_LWORD_TO_LREAL(bits);
      END_IF;
    END_IF;
  END_IF;
  was := x.DONE;
  IF x.DONE AND bad THEN
    DONE := FALSE;
    ERROR := TRUE;
    ERROR_ID := 7;
  END_IF;
END_FUNCTION_BLOCK

(* ---- CO_SDO_READ_STRING.st ---- *)
(*
 * CO_SDO_READ_STRING: reads object INDEX:SUBINDEX (a VISIBLE_STRING, up to
 * 254 characters before its first NUL) of node NODE (1..127) of CANopen
 * master network NETWORK into VALUE.
 * A rising edge of EXECUTE starts it; BUSY until the bridge has an answer,
 * then DONE or ERROR with ERROR_ID (docs/plc-library.md#sdo-blocks): 1 the
 * node aborted (ABORT_CODE), 2 no answer within TIMEOUT (T#0s: 5 s), 4 the
 * network is not running, 5 too many SDO requests wait, 6 invalid input,
 * 7 too large (more than 254 characters), 8 cancelled, 20 the bridge is not reachable, 22 the config
 * has no request mailbox.
 *)
(*
 * LINK is the generated `canworks.link` (ARRAY[0..1279] OF WORD); the block
 * uses a request mailbox of the bridge (`mailboxes` in the config, see
 * CW_LINK_SERVICE for the words). Instances share the request mailboxes in
 * the order they started.
 *)
FUNCTION_BLOCK CO_SDO_READ_STRING
VAR_INPUT
  EXECUTE : BOOL;
  NETWORK : USINT;
  NODE : USINT;
  INDEX : UINT;
  SUBINDEX : USINT;
  TIMEOUT : TIME;
END_VAR
VAR_OUTPUT
  BUSY : BOOL;
  DONE : BOOL;
  ERROR : BOOL;
  ERROR_ID : UINT;
  ABORT_CODE : UDINT;
  VALUE : STRING;
END_VAR
VAR_IN_OUT
  LINK : ARRAY[0..1279] OF WORD;
END_VAR
VAR
  x : CW_SDO_XFER;
  buf : ARRAY[0..1023] OF BYTE;
  was : BOOL;
  bad : BOOL;
  nchars : INT;
  i : INT;
END_VAR
  x(EXECUTE := EXECUTE, WRITE := FALSE, NETWORK := NETWORK, NODE := NODE, INDEX := INDEX, SUBINDEX := SUBINDEX,
    TIMEOUT := TIMEOUT, KIND := 2, MAX_SIZE := 16#FFFFFFFF, FETCH_MAX := 255, LINK := LINK, DATA := buf);
  BUSY := x.BUSY;
  DONE := x.DONE;
  ERROR := x.ERROR;
  ERROR_ID := x.ERROR_ID;
  ABORT_CODE := x.ABORT_CODE;
  IF x.DONE AND NOT was THEN
    nchars := UINT_TO_INT(x.GOT);
    FOR i := UINT_TO_INT(x.GOT) - 1 TO 0 BY -1 DO
      IF buf[i] = BYTE#0 THEN
        nchars := i;
      END_IF;
    END_FOR;
    bad := nchars > 254;
    IF NOT bad THEN
      VALUE := '';
      FOR i := 0 TO nchars - 1 DO
        VALUE := CONCAT(VALUE, CW_CHAR(buf[i]));
      END_FOR;
    END_IF;
  END_IF;
  was := x.DONE;
  IF x.DONE AND bad THEN
    DONE := FALSE;
    ERROR := TRUE;
    ERROR_ID := 7;
  END_IF;
END_FUNCTION_BLOCK

(* ---- CO_SDO_WRITE.st ---- *)
(*
 * CO_SDO_WRITE: writes DATA (SIZE 1 to 4 bytes, least significant first as
 * CANopen sends it) to object INDEX:SUBINDEX of node NODE (1..127) of
 * CANopen master network NETWORK, through the bridge's SDO registers; the
 * config needs "sdo_bridge_write": true.
 * A rising edge of EXECUTE starts it; BUSY until the bridge has an answer,
 * then DONE or ERROR with ERROR_ID (docs/plc-library.md): 1 the node aborted
 * (ABORT_CODE), 2 no answer within TIMEOUT (T#0s: 5 s), 6 invalid input,
 * 20 the bridge is not reachable, 21 SDO writes are not allowed by the
 * config (ABORT_CODE 16#08000020), 22 the config has no SDO registers,
 * 8 cancelled: the bridge restarted and did not send it (start it again).
 * Instances share the SDO registers: one waits while another uses them.
 *)
(*
 * LINK is the generated `canworks.link` (ARRAY[0..1279] OF WORD): the
 * bridge's blocks as canworks_in and canworks_out copy them from and to the
 * Modbus registers every scan, one word per register (high byte = the
 * bridge's even byte). Words: 0-3 status block, 4-6 control block, 7-13 SDO
 * request, 14-20 SDO response, 21 flags (bit 0 the bridge answers with this
 * program's map, 1 a control block, 2 SDO registers, 8 + n a live list for
 * network n), 22 control block owner, 23 SDO owner, 24 last instance number,
 * 25 + 8n .. 32 + 8n the live list of network n (n 0..7).
 *)
FUNCTION_BLOCK CO_SDO_WRITE
VAR_INPUT
  EXECUTE : BOOL;
  NETWORK : USINT;
  NODE : USINT;
  INDEX : UINT;
  SUBINDEX : USINT;
  DATA : UDINT;
  SIZE : USINT;
  TIMEOUT : TIME;
END_VAR
VAR_OUTPUT
  BUSY : BOOL;
  DONE : BOOL;
  ERROR : BOOL;
  ERROR_ID : UINT;
  ABORT_CODE : UDINT;
END_VAR
VAR_IN_OUT
  LINK : ARRAY[0..1279] OF WORD;
END_VAR
VAR
  me : WORD;
  prev : BOOL;
  phase : USINT;           (* 0 idle, 1 waiting for the SDO registers, 2 sent, 3 ended *)
  counter : WORD;
  timer : TON;
  state : WORD;
  err : UINT;
  fin : BOOL;
END_VAR
  IF me = WORD#0 THEN
    LINK[24] := UINT_TO_WORD(WORD_TO_UINT(LINK[24]) + 1);
    me := LINK[24];
  END_IF;
  IF phase = 3 AND NOT EXECUTE THEN
    phase := 0;
    DONE := FALSE;
    ERROR := FALSE;
  END_IF;
  err := 0;
  fin := FALSE;
  IF phase = 0 AND EXECUTE AND NOT prev THEN
    DONE := FALSE;
    ERROR := FALSE;
    ERROR_ID := 0;
    ABORT_CODE := 0;
    timer(IN := FALSE);
    IF (LINK[21] AND WORD#16#0001) = WORD#0 THEN
      err := 20;
    ELSIF (LINK[21] AND WORD#16#0004) = WORD#0 THEN
      err := 22;
    ELSIF NODE < 1 OR NODE > 127 OR SIZE < 1 OR SIZE > 4 THEN
      err := 6;
    ELSE
      phase := 1;
    END_IF;
  END_IF;
  IF phase = 1 OR phase = 2 THEN
    timer(IN := TRUE, PT := SEL(TIMEOUT = T#0s, TIMEOUT, T#5s));
    IF (LINK[21] AND WORD#16#0001) = WORD#0 THEN
      err := 20;
    ELSIF timer.Q THEN
      err := 2;
      ABORT_CODE := 16#05040000;
    ELSIF phase = 1 AND (LINK[23] = WORD#0 OR LINK[23] = me) THEN
      LINK[23] := me;
      counter := UINT_TO_WORD(WORD_TO_UINT(LINK[14]) + 1);
      LINK[7] := counter;
      LINK[8] := SHL(WORD#2, 8) OR USINT_TO_WORD(NETWORK);
      LINK[9] := SHL(USINT_TO_WORD(NODE), 8) OR USINT_TO_WORD(SUBINDEX);
      LINK[10] := UINT_TO_WORD(INDEX);
      LINK[11] := SHL(USINT_TO_WORD(SIZE), 8);
      LINK[12] := DWORD_TO_WORD(SHR(UDINT_TO_DWORD(DATA), 16));
      LINK[13] := DWORD_TO_WORD(UDINT_TO_DWORD(DATA));
      phase := 2;
    ELSIF phase = 2 AND LINK[14] = counter THEN
      state := SHR(LINK[15], 8);
      IF state = WORD#2 THEN
        fin := TRUE;
      ELSIF state = WORD#3 THEN
        ABORT_CODE := DWORD_TO_UDINT(SHL(WORD_TO_DWORD(LINK[16]), 16) OR WORD_TO_DWORD(LINK[17]));
        IF ABORT_CODE = 16#08000020 THEN
          err := 21;
        ELSIF ABORT_CODE = 16#08000021 THEN
          err := 8;            (* the bridge restarted and did not send it *)
        ELSE
          err := 1;
        END_IF;
      END_IF;
    END_IF;
  END_IF;
  IF err <> 0 OR fin THEN
    phase := 3;
    DONE := fin;
    ERROR := err <> 0;
    ERROR_ID := err;
    timer(IN := FALSE);
    IF LINK[23] = me THEN
      LINK[23] := WORD#0;
    END_IF;
  END_IF;
  BUSY := phase = 1 OR phase = 2;
  prev := EXECUTE;
END_FUNCTION_BLOCK

(* ---- CO_SDO_WRITE_BYTES.st ---- *)
(*
 * CO_SDO_WRITE_BYTES: writes the first SIZE bytes of BUFFER (up to 1024) to
 * object INDEX:SUBINDEX of node NODE (1..127) of CANopen master network
 * NETWORK, in one SDO download.
 * A rising edge of EXECUTE starts it; BUSY until the bridge has an answer,
 * then DONE or ERROR with ERROR_ID (docs/plc-library.md#sdo-blocks): 1 the
 * node aborted (ABORT_CODE), 2 no answer within TIMEOUT (T#0s: 5 s), 4 the
 * network is not running, 5 too many SDO requests wait, 6 invalid input,
 * 7 too large, 8 cancelled, 20 the bridge is not reachable, 22 the config
 * has no request mailbox.
 *)
(*
 * LINK is the generated `canworks.link` (ARRAY[0..1279] OF WORD); the block
 * uses a request mailbox of the bridge (`mailboxes` in the config, see
 * CW_LINK_SERVICE for the words). Instances share the request mailboxes in
 * the order they started.
 *)
FUNCTION_BLOCK CO_SDO_WRITE_BYTES
VAR_INPUT
  EXECUTE : BOOL;
  NETWORK : USINT;
  NODE : USINT;
  INDEX : UINT;
  SUBINDEX : USINT;
  TIMEOUT : TIME;
  SIZE : UINT;
END_VAR
VAR_OUTPUT
  BUSY : BOOL;
  DONE : BOOL;
  ERROR : BOOL;
  ERROR_ID : UINT;
  ABORT_CODE : UDINT;
END_VAR
VAR_IN_OUT
  BUFFER : ARRAY[0..1023] OF BYTE;
  LINK : ARRAY[0..1279] OF WORD;
END_VAR
VAR
  x : CW_SDO_XFER;
END_VAR
  x(EXECUTE := EXECUTE, WRITE := TRUE, NETWORK := NETWORK, NODE := NODE, INDEX := INDEX, SUBINDEX := SUBINDEX,
    TIMEOUT := TIMEOUT, KIND := 3, LENGTH := SIZE, LINK := LINK, DATA := BUFFER);
  BUSY := x.BUSY;
  DONE := x.DONE;
  ERROR := x.ERROR;
  ERROR_ID := x.ERROR_ID;
  ABORT_CODE := x.ABORT_CODE;
END_FUNCTION_BLOCK

(* ---- CO_SDO_WRITE_REAL.st ---- *)
(*
 * CO_SDO_WRITE_REAL: writes VALUE to object INDEX:SUBINDEX of node NODE
 * (1..127) of CANopen master network NETWORK, as REAL32 (SIZE 4), REAL64
 * (SIZE 8) or the object's type from its EDS (SIZE 0).
 * A rising edge of EXECUTE starts it; BUSY until the bridge has an answer,
 * then DONE or ERROR with ERROR_ID (docs/plc-library.md#sdo-blocks): 1 the
 * node aborted (ABORT_CODE), 2 no answer within TIMEOUT (T#0s: 5 s), 4 the
 * network is not running, 5 too many SDO requests wait, 6 invalid input,
 * 7 too large, 8 cancelled, 20 the bridge is not reachable, 22 the config
 * has no request mailbox.
 *)
(*
 * LINK is the generated `canworks.link` (ARRAY[0..1279] OF WORD); the block
 * uses a request mailbox of the bridge (`mailboxes` in the config, see
 * CW_LINK_SERVICE for the words). Instances share the request mailboxes in
 * the order they started.
 *)
FUNCTION_BLOCK CO_SDO_WRITE_REAL
VAR_INPUT
  EXECUTE : BOOL;
  NETWORK : USINT;
  NODE : USINT;
  INDEX : UINT;
  SUBINDEX : USINT;
  TIMEOUT : TIME;
  VALUE : LREAL;
  SIZE : USINT;
END_VAR
VAR_OUTPUT
  BUSY : BOOL;
  DONE : BOOL;
  ERROR : BOOL;
  ERROR_ID : UINT;
  ABORT_CODE : UDINT;
END_VAR
VAR_IN_OUT
  LINK : ARRAY[0..1279] OF WORD;
END_VAR
VAR
  x : CW_SDO_XFER;
  buf : ARRAY[0..1023] OF BYTE;
  prev : BOOL;
  bits : LWORD;
  i : INT;
END_VAR
  IF EXECUTE AND NOT prev AND NOT x.BUSY THEN
    bits := CW_LREAL_TO_LWORD(VALUE);
    FOR i := 0 TO 7 DO
      buf[i] := LWORD_TO_BYTE(SHR(bits, 8 * i));
    END_FOR;
  END_IF;
  prev := EXECUTE;
  x(EXECUTE := EXECUTE, WRITE := TRUE, NETWORK := NETWORK, NODE := NODE, INDEX := INDEX, SUBINDEX := SUBINDEX,
    TIMEOUT := TIMEOUT, KIND := 1, SIZE := SIZE, LENGTH := 8, LINK := LINK, DATA := buf);
  BUSY := x.BUSY;
  DONE := x.DONE;
  ERROR := x.ERROR;
  ERROR_ID := x.ERROR_ID;
  ABORT_CODE := x.ABORT_CODE;
END_FUNCTION_BLOCK

(* ---- CO_SDO_WRITE_STRING.st ---- *)
(*
 * CO_SDO_WRITE_STRING: writes VALUE (its characters, up to 254, without a
 * NUL) to object INDEX:SUBINDEX of node NODE (1..127) of CANopen master
 * network NETWORK.
 * A rising edge of EXECUTE starts it; BUSY until the bridge has an answer,
 * then DONE or ERROR with ERROR_ID (docs/plc-library.md#sdo-blocks): 1 the
 * node aborted (ABORT_CODE), 2 no answer within TIMEOUT (T#0s: 5 s), 4 the
 * network is not running, 5 too many SDO requests wait, 6 invalid input,
 * 7 too large, 8 cancelled, 20 the bridge is not reachable, 22 the config
 * has no request mailbox.
 *)
(*
 * LINK is the generated `canworks.link` (ARRAY[0..1279] OF WORD); the block
 * uses a request mailbox of the bridge (`mailboxes` in the config, see
 * CW_LINK_SERVICE for the words). Instances share the request mailboxes in
 * the order they started.
 *)
FUNCTION_BLOCK CO_SDO_WRITE_STRING
VAR_INPUT
  EXECUTE : BOOL;
  NETWORK : USINT;
  NODE : USINT;
  INDEX : UINT;
  SUBINDEX : USINT;
  TIMEOUT : TIME;
  VALUE : STRING;
END_VAR
VAR_OUTPUT
  BUSY : BOOL;
  DONE : BOOL;
  ERROR : BOOL;
  ERROR_ID : UINT;
  ABORT_CODE : UDINT;
END_VAR
VAR_IN_OUT
  LINK : ARRAY[0..1279] OF WORD;
END_VAR
VAR
  x : CW_SDO_XFER;
  buf : ARRAY[0..1023] OF BYTE;
  prev : BOOL;
  nchars : INT;
  i : INT;
END_VAR
  IF EXECUTE AND NOT prev AND NOT x.BUSY THEN
    nchars := LEN(VALUE);
    IF nchars > 254 THEN
      nchars := 254;
    END_IF;
    FOR i := 1 TO nchars DO
      buf[i - 1] := CW_CHAR_CODE(MID(VALUE, 1, i));
    END_FOR;
  END_IF;
  prev := EXECUTE;
  x(EXECUTE := EXECUTE, WRITE := TRUE, NETWORK := NETWORK, NODE := NODE, INDEX := INDEX, SUBINDEX := SUBINDEX,
    TIMEOUT := TIMEOUT, KIND := 2, LENGTH := INT_TO_UINT(nchars), LINK := LINK, DATA := buf);
  BUSY := x.BUSY;
  DONE := x.DONE;
  ERROR := x.ERROR;
  ERROR_ID := x.ERROR_ID;
  ABORT_CODE := x.ABORT_CODE;
END_FUNCTION_BLOCK

(* ---- CW_LINK_SERVICE.st ---- *)
(*
 * CW_LINK_SERVICE: the start of every scan for the blocks that use the
 * bridge's mailboxes (bridge-plc-blocks). The generated canworks_in calls it
 * once, after it copied the input words into LINK and before any user code:
 * it counts the scan, moves the lowest waiting mailbox ticket of the last
 * scan into place, frees a request mailbox whose owner was not called for
 * 100 scans and marks the receivers of a new receive batch pending. While
 * the bridge is not reachable it clears the requests and the
 * acknowledgement, so that a restarted bridge never runs an old request.
 *)
(*
 * The mailbox words of LINK (ARRAY[0..1279] OF WORD), after change 1's 0-88:
 * 89 flags (bits 0-2 request mailboxes, 4 receive mailbox, 5 network info,
 * 8-12 cyclic jobs), 90 scan counter, 91 last ticket, 92 lowest ticket
 * waiting in this scan, 93 the same of the last scan, 94-97 mailbox owners,
 * 98-101 owner stamps (scan counter), 102 receive batch seen, 103-104 the
 * receivers still pending (word 103 bits 31-16), 105 last batch taken,
 * 128 + j keepalive of cyclic job j, 144 + 144m request mailbox m (72
 * request words, then 72 response words), 720 the receive mailbox (120
 * words per receive block, 2 at most), 960 + 18n the info of network n, 1104
 * the cyclic job table.
 *)
FUNCTION_BLOCK CW_LINK_SERVICE
VAR_IN_OUT
  LINK : ARRAY[0..1279] OF WORD;
END_VAR
VAR
  m : INT;
END_VAR
  LINK[90] := UDINT_TO_WORD(WORD_TO_UDINT(LINK[90]) + 1);
  LINK[93] := LINK[92];
  LINK[92] := WORD#0;
  IF (LINK[21] AND WORD#16#0001) = WORD#0 THEN
    FOR m := 0 TO 3 DO
      LINK[144 + 144 * m + 1] := WORD#0;
      LINK[94 + m] := WORD#0;
    END_FOR;
    LINK[102] := WORD#0;
    LINK[103] := WORD#0;
    LINK[104] := WORD#0;
    LINK[105] := WORD#0;
    RETURN;
  END_IF;
  FOR m := 0 TO 3 DO
    IF LINK[94 + m] <> WORD#0 AND DINT_TO_WORD(WORD_TO_DINT(LINK[90]) - WORD_TO_DINT(LINK[98 + m])) > WORD#100 THEN
      LINK[94 + m] := WORD#0;
    END_IF;
  END_FOR;
  IF (LINK[89] AND WORD#16#0010) <> WORD#0 AND LINK[720] <> LINK[105] THEN
    LINK[105] := LINK[720];
    LINK[102] := LINK[720];
    LINK[103] := LINK[721];
    LINK[104] := LINK[722];
  END_IF;
END_FUNCTION_BLOCK

(* ---- CW_MB_CALL.st ---- *)
(*
 * CW_MB_CALL: one block's use of a request mailbox of the bridge
 * (bridge-plc-blocks), for the blocks of this library.
 * While RUN is TRUE it waits for a free mailbox in ticket order (the
 * waiting instance with the lowest ticket of the last scan goes first),
 * then keeps it (OWNED, request words from LINK[BASE], response words from
 * LINK[BASE + 72]) and stamps it every call. A call with SEND while OWNED and
 * not WAITING writes the request: OP, NET, A0..A5; the caller puts the data
 * words at LINK[BASE + 8] first. ANSWERED is TRUE in the call that sees the
 * answer, with ERR its ERROR_ID (0: done); the results are at LINK[BASE + 74]
 * and the data at LINK[BASE + 80]. RUN FALSE frees the mailbox. LOST: the
 * bridge is not reachable (the block ends with ERROR_ID 20); the mailbox is
 * freed.
 *)
FUNCTION_BLOCK CW_MB_CALL
VAR_INPUT
  RUN : BOOL;
  SEND : BOOL;
  OP : USINT;
  NET : USINT;
  A0 : WORD;
  A1 : WORD;
  A2 : WORD;
  A3 : WORD;
  A4 : WORD;
  A5 : WORD;
END_VAR
VAR_OUTPUT
  OWNED : BOOL;
  BASE : INT;
  WAITING : BOOL;
  ANSWERED : BOOL;
  ERR : UINT;
  LOST : BOOL;
END_VAR
VAR_IN_OUT
  LINK : ARRAY[0..1279] OF WORD;
END_VAR
VAR
  me : WORD;
  ticket : WORD;
  m : INT;
  i : INT;
  cnt : INT;
  counter : WORD;
END_VAR
  IF me = WORD#0 THEN
    LINK[24] := UDINT_TO_WORD(WORD_TO_UDINT(LINK[24]) + 1);
    me := LINK[24];
  END_IF;
  ANSWERED := FALSE;
  LOST := (LINK[21] AND WORD#16#0001) = WORD#0;
  IF OWNED AND LINK[94 + m] <> me THEN
    LOST := TRUE;
    OWNED := FALSE;
  END_IF;
  IF NOT RUN OR LOST THEN
    IF OWNED AND LINK[94 + m] = me THEN
      LINK[94 + m] := WORD#0;
    END_IF;
    OWNED := FALSE;
    WAITING := FALSE;
    ticket := WORD#0;
    RETURN;
  END_IF;
  IF NOT OWNED THEN
    IF ticket = WORD#0 THEN
      LINK[91] := UDINT_TO_WORD(WORD_TO_UDINT(LINK[91]) + 1);
      IF LINK[91] = WORD#0 THEN
        LINK[91] := WORD#1;
      END_IF;
      ticket := LINK[91];
    END_IF;
    cnt := WORD_TO_INT(LINK[89] AND WORD#16#0007);
    IF cnt > 4 THEN
      cnt := 4;
    END_IF;
    (* My turn: nobody waited in the last scan, or I was the lowest. *)
    IF LINK[93] = WORD#0 OR ticket = LINK[93] OR (DINT_TO_WORD(WORD_TO_DINT(ticket) - WORD_TO_DINT(LINK[93])) AND WORD#16#8000) <> WORD#0 THEN
      FOR i := 0 TO cnt - 1 DO
        IF NOT OWNED AND LINK[94 + i] = WORD#0 THEN
          m := i;
          OWNED := TRUE;
        END_IF;
      END_FOR;
    END_IF;
    IF OWNED THEN
      LINK[94 + m] := me;
      BASE := 144 + 144 * m;
      WAITING := FALSE;
      ticket := WORD#0;
    ELSIF LINK[92] = WORD#0 OR (DINT_TO_WORD(WORD_TO_DINT(ticket) - WORD_TO_DINT(LINK[92])) AND WORD#16#8000) <> WORD#0 THEN
      LINK[92] := ticket;
    END_IF;
  END_IF;
  IF NOT OWNED THEN
    RETURN;
  END_IF;
  LINK[98 + m] := LINK[90];
  IF SEND AND NOT WAITING THEN
    (* A counter the bridge has not seen: not the last request, not the echo. *)
    counter := UDINT_TO_WORD(WORD_TO_UDINT(LINK[BASE]) + 1);
    IF counter = LINK[BASE + 72] THEN
      counter := UDINT_TO_WORD(WORD_TO_UDINT(counter) + 1);
    END_IF;
    LINK[BASE] := counter;
    LINK[BASE + 1] := SHL(USINT_TO_WORD(OP), 8) OR USINT_TO_WORD(NET);
    LINK[BASE + 2] := A0;
    LINK[BASE + 3] := A1;
    LINK[BASE + 4] := A2;
    LINK[BASE + 5] := A3;
    LINK[BASE + 6] := A4;
    LINK[BASE + 7] := A5;
    WAITING := TRUE;
  ELSIF WAITING AND LINK[BASE + 72] = counter AND SHR(LINK[BASE + 73], 8) >= WORD#2 THEN
    WAITING := FALSE;
    ANSWERED := TRUE;
    ERR := WORD_TO_UINT(LINK[BASE + 73] AND WORD#16#00FF);
  END_IF;
END_FUNCTION_BLOCK

(* ---- CW_REQUEST.st ---- *)
(*
 * CW_REQUEST: one operation through a request mailbox of the bridge, for
 * the CAN and J1939 blocks of this library. A rising edge of EXECUTE starts
 * it: the first LENGTH bytes of DATA go with it (more than 128 go to the
 * bridge first with STAGE requests), then OP on network NET with arguments
 * A0..A5. The answer's results are R0..R5; with RLEN_AT 0..5 that result is
 * the length of the answer's data, which is fetched into DATA (FETCH
 * requests after the first 128 bytes, at most FETCH_MAX); with RLEN_AT 6,
 * FETCH_MAX bytes of the first part are copied. ERROR_ID: the bridge's, or
 * 20 the bridge is not reachable, 22 the config has no request mailbox.
 *)
FUNCTION_BLOCK CW_REQUEST
VAR_INPUT
  EXECUTE : BOOL;
  OP : USINT;
  NET : USINT;
  A0 : WORD;
  A1 : WORD;
  A2 : WORD;
  A3 : WORD;
  A4 : WORD;
  A5 : WORD;
  LENGTH : UINT;
  RLEN_AT : INT := 6;
  FETCH_MAX : UINT;
END_VAR
VAR_OUTPUT
  BUSY : BOOL;
  DONE : BOOL;
  ERROR : BOOL;
  ERROR_ID : UINT;
  R0 : WORD;
  R1 : WORD;
  R2 : WORD;
  R3 : WORD;
  R4 : WORD;
  R5 : WORD;
  GOT : UINT;
END_VAR
VAR_IN_OUT
  LINK : ARRAY[0..1279] OF WORD;
  DATA : ARRAY[0..1784] OF BYTE;
END_VAR
VAR
  mb : CW_MB_CALL;
  prev : BOOL;
  phase : USINT;           (* 0 idle, 1 staging, 2 the operation, 3 fetching, 4 ended *)
  offset : UINT;
  want : UINT;
  cnt : INT;
  k : INT;
  b : INT;
  err : UINT;
  fin : BOOL;
  rlen : WORD;
END_VAR
  IF phase = 4 AND NOT EXECUTE THEN
    phase := 0;
    DONE := FALSE;
    ERROR := FALSE;
  END_IF;
  err := 0;
  fin := FALSE;
  IF phase = 0 AND EXECUTE AND NOT prev THEN
    DONE := FALSE;
    ERROR := FALSE;
    ERROR_ID := 0;
    GOT := 0;
    offset := 0;
    IF (LINK[21] AND WORD#16#0001) = WORD#0 THEN
      err := 20;
    ELSIF (LINK[89] AND WORD#16#0007) = WORD#0 THEN
      err := 22;
    ELSIF LENGTH > 128 THEN
      phase := 1;
    ELSE
      phase := 2;
    END_IF;
  END_IF;
  IF phase >= 1 AND phase <= 3 THEN
    mb(RUN := TRUE, SEND := FALSE, LINK := LINK);
    b := mb.BASE;
    IF mb.LOST THEN
      err := 20;
    ELSIF mb.ANSWERED AND mb.ERR <> 0 THEN
      err := mb.ERR;
      IF phase = 2 THEN
        R0 := LINK[b + 74];
        R1 := LINK[b + 75];
        R2 := LINK[b + 76];
        R3 := LINK[b + 77];
        R4 := LINK[b + 78];
        R5 := LINK[b + 79];
      END_IF;
    ELSIF mb.ANSWERED AND phase = 1 THEN
      offset := offset + 128;
      IF offset >= LENGTH THEN
        phase := 2;
      END_IF;
    ELSIF mb.ANSWERED THEN
      IF phase = 2 THEN
        R0 := LINK[b + 74];
        R1 := LINK[b + 75];
        R2 := LINK[b + 76];
        R3 := LINK[b + 77];
        R4 := LINK[b + 78];
        R5 := LINK[b + 79];
        want := FETCH_MAX;
        IF RLEN_AT >= 0 AND RLEN_AT <= 5 THEN
          rlen := LINK[b + 74 + RLEN_AT];
          IF WORD_TO_UINT(rlen) < want THEN
            want := WORD_TO_UINT(rlen);
          END_IF;
        ELSIF want > 128 THEN
          want := 128;
        END_IF;
        IF want > 1785 THEN
          want := 1785;
        END_IF;
      END_IF;
      cnt := UINT_TO_INT(want - GOT);
      IF cnt > 128 THEN
        cnt := 128;
      END_IF;
      FOR k := 0 TO cnt - 1 DO
        IF (k MOD 2) = 0 THEN
          DATA[UINT_TO_INT(GOT) + k] := WORD_TO_BYTE(SHR(LINK[b + 80 + k / 2], 8));
        ELSE
          DATA[UINT_TO_INT(GOT) + k] := WORD_TO_BYTE(LINK[b + 80 + k / 2]);
        END_IF;
      END_FOR;
      GOT := GOT + INT_TO_UINT(cnt);
      IF GOT >= want THEN
        fin := TRUE;
      ELSE
        phase := 3;
      END_IF;
    END_IF;
    IF err = 0 AND NOT fin AND mb.OWNED AND NOT mb.WAITING THEN
      IF phase = 1 OR (phase = 2 AND LENGTH <= 128) THEN
        cnt := UINT_TO_INT(LENGTH - offset);
        IF cnt > 128 THEN
          cnt := 128;
        END_IF;
        FOR k := 0 TO 63 DO
          LINK[b + 8 + k] := WORD#0;
        END_FOR;
        FOR k := 0 TO cnt - 1 DO
          IF (k MOD 2) = 0 THEN
            LINK[b + 8 + k / 2] := SHL(BYTE_TO_WORD(DATA[UINT_TO_INT(offset) + k]), 8);
          ELSE
            LINK[b + 8 + k / 2] := LINK[b + 8 + k / 2] OR BYTE_TO_WORD(DATA[UINT_TO_INT(offset) + k]);
          END_IF;
        END_FOR;
      END_IF;
      IF phase = 1 THEN
        mb(RUN := TRUE, SEND := TRUE, OP := 1, NET := 0, A0 := UINT_TO_WORD(offset), A1 := INT_TO_WORD(cnt),
           A2 := WORD#0, A3 := WORD#0, A4 := WORD#0, A5 := WORD#0, LINK := LINK);
      ELSIF phase = 2 THEN
        mb(RUN := TRUE, SEND := TRUE, OP := OP, NET := NET, A0 := A0, A1 := A1, A2 := A2, A3 := A3, A4 := A4,
           A5 := A5, LINK := LINK);
      ELSE
        mb(RUN := TRUE, SEND := TRUE, OP := 2, NET := 0, A0 := UINT_TO_WORD(GOT), A1 := WORD#0, A2 := WORD#0, A3 := WORD#0,
           A4 := WORD#0, A5 := WORD#0, LINK := LINK);
      END_IF;
    END_IF;
  END_IF;
  IF err <> 0 OR fin THEN
    phase := 4;
    DONE := fin;
    ERROR := err <> 0;
    ERROR_ID := err;
    mb(RUN := FALSE, LINK := LINK);
  END_IF;
  BUSY := phase >= 1 AND phase <= 3;
  prev := EXECUTE;
END_FUNCTION_BLOCK

(* ---- CW_RX.st ---- *)
(*
 * CW_RX: one receiver of the bridge's receive mailbox, for the receiving
 * blocks of this library (CAN_RECEIVE, J1939_RECEIVE, CO_RECV_EMCY).
 * While ENABLE is TRUE it keeps a receiver of KIND (1 CAN, 2 J1939, 3 EMCY)
 * open with FLAGS, DEPTH, ID and MASK (RX_OPEN through a request mailbox);
 * CHANGED closes it and opens it again. A call with NEXT delivers the next
 * record of this receiver in the current batch: RECEIVED, its first word at
 * LINK[REC]. When the batch has no more of them the receiver's pending mark
 * is cleared, so the bridge can show the next batch. After an error whose
 * bit is set in RETRY (bit n for ERROR_ID n) it opens the receiver again on
 * the next call; 8 means the bridge closed it (link stop, stall, network
 * restart). ENABLE FALSE closes it (RX_CLOSE).
 *)
FUNCTION_BLOCK CW_RX
VAR_INPUT
  ENABLE : BOOL;
  CHANGED : BOOL;
  NEXT : BOOL;
  KIND : USINT;
  NETWORK : USINT;
  FLAGS : USINT;
  DEPTH : UINT;
  ID : UDINT;
  MASK : UDINT;
  RETRY : DWORD;
END_VAR
VAR_OUTPUT
  ACTIVE : BOOL;
  RECEIVED : BOOL;
  REC : INT;
  ERROR : BOOL;
  ERROR_ID : UINT;
  SLOT : INT;
END_VAR
VAR_IN_OUT
  LINK : ARRAY[0..1279] OF WORD;
END_VAR
VAR
  mb : CW_MB_CALL;
  prev : BOOL;
  phase : USINT;           (* 0 closed, 1 opening, 2 open, 3 closing *)
  gen : WORD;
  tick0 : WORD;
  seq : WORD;
  pos : INT;
  pw : INT;
  slot_bit : WORD;
  shown : WORD;
  hdr : WORD;
  size : INT;
  synced : BOOL;          (* the batch on show was built after the open *)
  fresh : BOOL;
  found : BOOL;
  err : UINT;
END_VAR
  RECEIVED := FALSE;
  err := 0;
  IF ENABLE AND NOT prev THEN
    ERROR := FALSE;
    ERROR_ID := 0;
  END_IF;
  IF (LINK[21] AND WORD#16#0001) = WORD#0 AND phase <> 0 THEN
    (* The bridge ended every receiver when the link stopped. *)
    mb(RUN := FALSE, LINK := LINK);
    phase := 0;
    IF ENABLE THEN
      err := 20;
    END_IF;
  END_IF;
  IF phase = 2 THEN
    IF NOT synced THEN
      synced := (DINT_TO_WORD(WORD_TO_DINT(LINK[724]) - WORD_TO_DINT(tick0)) AND WORD#16#8000) = WORD#0;
    END_IF;
    fresh := synced;
    shown := SHR(LINK[725 + SLOT / 2], 8 * (1 - SLOT MOD 2)) AND WORD#16#00FF;
    IF fresh AND shown <> gen THEN
      phase := 0;
      err := 8;
    ELSIF NOT ENABLE OR CHANGED THEN
      phase := 3;
    END_IF;
  END_IF;
  IF phase = 2 OR phase = 3 THEN
    pw := 104 - SLOT / 16;
    slot_bit := SHL(WORD#1, SLOT MOD 16);
  END_IF;
  IF phase = 3 THEN
    LINK[pw] := LINK[pw] AND NOT slot_bit;
  END_IF;
  IF phase = 0 AND ENABLE AND err = 0 AND
     NOT (ERROR AND (SHR(RETRY, UINT_TO_INT(ERROR_ID)) AND DWORD#16#00000001) = DWORD#0) THEN
    ERROR := FALSE;
    ERROR_ID := 0;
    IF (LINK[21] AND WORD#16#0001) = WORD#0 THEN
      err := 20;
    ELSIF (LINK[89] AND WORD#16#0007) = WORD#0 OR (LINK[89] AND WORD#16#0010) = WORD#0 THEN
      err := 22;
    ELSE
      phase := 1;
    END_IF;
  END_IF;
  IF phase = 1 OR phase = 3 THEN
    mb(RUN := TRUE, SEND := FALSE, LINK := LINK);
    IF mb.LOST THEN
      phase := 0;
      err := SEL(ENABLE, UINT#0, UINT#20);
    ELSIF mb.ANSWERED AND phase = 1 THEN
      IF mb.ERR <> 0 THEN
        err := mb.ERR;
        phase := 0;
      ELSE
        SLOT := WORD_TO_INT(LINK[mb.BASE + 74]);
        gen := LINK[mb.BASE + 75];
        tick0 := LINK[mb.BASE + 76];
        synced := FALSE;
        seq := WORD#0;
        pos := 0;
        phase := 2;
      END_IF;
      mb(RUN := FALSE, LINK := LINK);
    ELSIF mb.ANSWERED THEN
      phase := 0;
      mb(RUN := FALSE, LINK := LINK);
    ELSIF mb.OWNED AND NOT mb.WAITING THEN
      IF phase = 1 THEN
        mb(RUN := TRUE, SEND := TRUE, OP := 8, NET := NETWORK,
           A0 := SHL(USINT_TO_WORD(KIND), 8) OR USINT_TO_WORD(FLAGS), A1 := UINT_TO_WORD(DEPTH),
           A2 := DWORD_TO_WORD(SHR(UDINT_TO_DWORD(ID), 16)), A3 := UDINT_TO_WORD(ID),
           A4 := DWORD_TO_WORD(SHR(UDINT_TO_DWORD(MASK), 16)), A5 := UDINT_TO_WORD(MASK), LINK := LINK);
      ELSE
        mb(RUN := TRUE, SEND := TRUE, OP := 9, NET := NETWORK, A0 := INT_TO_WORD(SLOT), A1 := WORD#0, A2 := WORD#0, A3 := WORD#0,
           A4 := WORD#0, A5 := WORD#0, LINK := LINK);
      END_IF;
    END_IF;
  END_IF;
  IF phase = 2 AND NEXT THEN
    (* My records of the batch on show: only in a batch built after the open
       (its present slot_bit set while the block is newer than the open) and while
       still pending. *)
    pw := 104 - SLOT / 16;
    slot_bit := SHL(WORD#1, SLOT MOD 16);
    IF LINK[720] <> seq THEN
      seq := LINK[720];
      pos := 745;
    END_IF;
    IF NOT synced THEN
      synced := (DINT_TO_WORD(WORD_TO_DINT(LINK[724]) - WORD_TO_DINT(tick0)) AND WORD#16#8000) = WORD#0;
    END_IF;
    fresh := synced;
    IF fresh AND (LINK[722 - SLOT / 16] AND slot_bit) <> WORD#0 AND (LINK[pw] AND slot_bit) <> WORD#0 THEN
      found := FALSE;
      WHILE NOT found AND pos < 745 + WORD_TO_INT(LINK[723]) AND pos < 960 DO
        hdr := LINK[pos];
        size := 7;
        CASE WORD_TO_INT(SHR(hdr, 4) AND WORD#16#000F) OF
          1: size := 10;
          2: size := 12;
          3: size := 12;
        END_CASE;
        IF WORD_TO_INT(SHR(hdr, 8)) = SLOT THEN
          found := TRUE;
          REC := pos;
          RECEIVED := TRUE;
        END_IF;
        pos := pos + size;
      END_WHILE;
      IF NOT found THEN
        LINK[pw] := LINK[pw] AND NOT slot_bit;
      END_IF;
    END_IF;
  END_IF;
  IF err <> 0 THEN
    ERROR := TRUE;
    ERROR_ID := err;
  END_IF;
  ACTIVE := phase = 2;
  prev := ENABLE;
END_FUNCTION_BLOCK

(* ---- CW_SDO_XFER.st ---- *)
(*
 * CW_SDO_XFER: one SDO transfer through a request mailbox of the bridge,
 * for the SDO blocks of this library (CO_SDO_READ_BYTES and the others).
 * A rising edge of EXECUTE starts it. A write sends LENGTH bytes of DATA
 * (more than 128 go to the bridge first with STAGE requests); a read
 * answers RSIZE, the object's size, and fetches its first
 * MIN(RSIZE, FETCH_MAX, 1024) bytes into DATA (FETCH requests after the
 * first 128). KIND: 1 REAL, 2 STRING, 3 bytes; SIZE the REAL write's size.
 * ERROR_IDs as the bridge gives them (docs/plc-library.md#sdo-blocks) and
 * 6 invalid input, 7 a reply longer than MAX_SIZE, 20 the bridge is not
 * reachable, 22 the config has no request mailbox.
 *)
FUNCTION_BLOCK CW_SDO_XFER
VAR_INPUT
  EXECUTE : BOOL;
  WRITE : BOOL;
  NETWORK : USINT;
  NODE : USINT;
  INDEX : UINT;
  SUBINDEX : USINT;
  TIMEOUT : TIME;
  KIND : USINT;
  SIZE : USINT;
  LENGTH : UINT;
  MAX_SIZE : UDINT := 1024;
  FETCH_MAX : UINT := 1024;
END_VAR
VAR_OUTPUT
  BUSY : BOOL;
  DONE : BOOL;
  ERROR : BOOL;
  ERROR_ID : UINT;
  ABORT_CODE : UDINT;
  RSIZE : UDINT;
  GOT : UINT;
END_VAR
VAR_IN_OUT
  LINK : ARRAY[0..1279] OF WORD;
  DATA : ARRAY[0..1023] OF BYTE;
END_VAR
VAR
  mb : CW_MB_CALL;
  prev : BOOL;
  phase : USINT;           (* 0 idle, 1 staging, 2 the operation, 3 fetching, 4 ended *)
  offset : UINT;
  want : UINT;
  cnt : INT;
  k : INT;
  b : INT;
  ms : UDINT;
  err : UINT;
  fin : BOOL;
  op : USINT;
END_VAR
  IF phase = 4 AND NOT EXECUTE THEN
    phase := 0;
    DONE := FALSE;
    ERROR := FALSE;
  END_IF;
  err := 0;
  fin := FALSE;
  IF phase = 0 AND EXECUTE AND NOT prev THEN
    DONE := FALSE;
    ERROR := FALSE;
    ERROR_ID := 0;
    ABORT_CODE := 0;
    RSIZE := 0;
    GOT := 0;
    offset := 0;
    IF (LINK[21] AND WORD#16#0001) = WORD#0 THEN
      err := 20;
    ELSIF (LINK[89] AND WORD#16#0007) = WORD#0 THEN
      err := 22;
    ELSIF NODE < 1 OR NODE > 127 OR (WRITE AND LENGTH > 1024) THEN
      err := 6;
    ELSIF WRITE AND LENGTH > 128 THEN
      phase := 1;
    ELSE
      phase := 2;
    END_IF;
  END_IF;
  IF phase >= 1 AND phase <= 3 THEN
    mb(RUN := TRUE, SEND := FALSE, LINK := LINK);
    b := mb.BASE;
    IF mb.LOST THEN
      err := 20;
    ELSIF mb.ANSWERED AND mb.ERR <> 0 THEN
      err := mb.ERR;
      IF phase = 2 THEN
        ABORT_CODE := WORD_TO_UDINT(LINK[b + 76]) * 65536 + WORD_TO_UDINT(LINK[b + 77]);
      END_IF;
    ELSIF mb.ANSWERED AND phase = 1 THEN
      offset := offset + 128;
      IF offset >= LENGTH THEN
        phase := 2;
      END_IF;
    ELSIF mb.ANSWERED AND phase = 2 AND WRITE THEN
      fin := TRUE;
    ELSIF mb.ANSWERED THEN
      IF phase = 2 THEN
        RSIZE := WORD_TO_UDINT(LINK[b + 74]) * 65536 + WORD_TO_UDINT(LINK[b + 75]);
        want := FETCH_MAX;
        IF want > 1024 THEN
          want := 1024;
        END_IF;
        IF RSIZE < UINT_TO_UDINT(want) THEN
          want := UDINT_TO_UINT(RSIZE);
        END_IF;
      END_IF;
      IF phase = 2 AND RSIZE > MAX_SIZE THEN
        err := 7;
      ELSE
        cnt := UINT_TO_INT(want - GOT);
        IF cnt > 128 THEN
          cnt := 128;
        END_IF;
        FOR k := 0 TO cnt - 1 DO
          IF (k MOD 2) = 0 THEN
            DATA[UINT_TO_INT(GOT) + k] := WORD_TO_BYTE(SHR(LINK[b + 80 + k / 2], 8));
          ELSE
            DATA[UINT_TO_INT(GOT) + k] := WORD_TO_BYTE(LINK[b + 80 + k / 2]);
          END_IF;
        END_FOR;
        GOT := GOT + INT_TO_UINT(cnt);
        IF GOT >= want THEN
          fin := TRUE;
        ELSE
          phase := 3;
        END_IF;
      END_IF;
    END_IF;
    IF err = 0 AND NOT fin AND mb.OWNED AND NOT mb.WAITING THEN
      IF phase = 1 THEN
        cnt := UINT_TO_INT(LENGTH - offset);
        IF cnt > 128 THEN
          cnt := 128;
        END_IF;
        FOR k := 0 TO 63 DO
          LINK[b + 8 + k] := WORD#0;
        END_FOR;
        FOR k := 0 TO cnt - 1 DO
          IF (k MOD 2) = 0 THEN
            LINK[b + 8 + k / 2] := SHL(BYTE_TO_WORD(DATA[UINT_TO_INT(offset) + k]), 8);
          ELSE
            LINK[b + 8 + k / 2] := LINK[b + 8 + k / 2] OR BYTE_TO_WORD(DATA[UINT_TO_INT(offset) + k]);
          END_IF;
        END_FOR;
        mb(RUN := TRUE, SEND := TRUE, OP := 1, NET := 0, A0 := UINT_TO_WORD(offset), A1 := INT_TO_WORD(cnt),
           A2 := WORD#0, A3 := WORD#0, A4 := WORD#0, A5 := WORD#0, LINK := LINK);
      ELSIF phase = 2 THEN
        IF WRITE AND LENGTH <= 128 THEN
          FOR k := 0 TO 63 DO
            LINK[b + 8 + k] := WORD#0;
          END_FOR;
          FOR k := 0 TO UINT_TO_INT(LENGTH) - 1 DO
            IF (k MOD 2) = 0 THEN
              LINK[b + 8 + k / 2] := SHL(BYTE_TO_WORD(DATA[k]), 8);
            ELSE
              LINK[b + 8 + k / 2] := LINK[b + 8 + k / 2] OR BYTE_TO_WORD(DATA[k]);
            END_IF;
          END_FOR;
        END_IF;
        ms := DWORD_TO_UDINT(TIME_TO_DWORD(TIMEOUT));
        IF ms > 65535 THEN
          ms := 65535;
        END_IF;
        op := SEL(WRITE, USINT#3, USINT#4);
        mb(RUN := TRUE, SEND := TRUE, OP := op, NET := NETWORK,
           A0 := SHL(USINT_TO_WORD(NODE), 8) OR USINT_TO_WORD(SUBINDEX), A1 := UINT_TO_WORD(INDEX),
           A2 := SHL(USINT_TO_WORD(KIND), 8) OR USINT_TO_WORD(SIZE), A3 := UDINT_TO_WORD(ms),
           A4 := UINT_TO_WORD(LENGTH), A5 := WORD#0, LINK := LINK);
      ELSE
        mb(RUN := TRUE, SEND := TRUE, OP := 2, NET := 0, A0 := UINT_TO_WORD(GOT), A1 := WORD#0, A2 := WORD#0, A3 := WORD#0,
           A4 := WORD#0, A5 := WORD#0, LINK := LINK);
      END_IF;
    END_IF;
  END_IF;
  IF err <> 0 OR fin THEN
    phase := 4;
    DONE := fin;
    ERROR := err <> 0;
    ERROR_ID := err;
    mb(RUN := FALSE, LINK := LINK);
  END_IF;
  BUSY := phase >= 1 AND phase <= 3;
  prev := EXECUTE;
END_FUNCTION_BLOCK

(* ---- J1939_DM_CLEAR.st ---- *)
(*
 * J1939_DM_CLEAR: clears the trouble codes of ECU DESTINATION (255: every
 * ECU) on J1939 network NETWORK: the previously active ones (DM3,
 * PREVIOUS_ONLY) or the active and previously active ones (DM11). A rising edge of EXECUTE starts it; BUSY until the bridge has
 * an answer, then DONE or ERROR with ERROR_ID (docs/plc-library.md#j1939-blocks):
 * 1 the network is not running, 2 no such network, 3 invalid input,
 * 4 the network sends that PGN itself, 5 another DM2 read or clear for that
 * address is pending, 6 no answer within TIMEOUT, 7 the bus is off,
 * 8 cancelled, 9 no free job or receiver, 10 not a J1939 network, 11 the
 * network holds no address, 12 the destination answered NACK, 13 no DM1
 * from that source, 14 the transfer was aborted, 20 the bridge is not
 * reachable, 22 the config has no request mailbox.
 *)
(*
 * LINK is the generated `canworks.link` (ARRAY[0..1279] OF WORD); the block uses a request mailbox of the bridge (`mailboxes` in the config); instances share
 * them in the order they started (see
 * CW_LINK_SERVICE for the words).
 *)
FUNCTION_BLOCK J1939_DM_CLEAR
VAR_INPUT
  EXECUTE : BOOL;
  NETWORK : USINT;
  DESTINATION : USINT;
  PREVIOUS_ONLY : BOOL;
  TIMEOUT : TIME;
END_VAR
VAR_IN_OUT
  LINK : ARRAY[0..1279] OF WORD;
END_VAR
VAR_OUTPUT
  BUSY : BOOL;
  DONE : BOOL;
  ERROR : BOOL;
  ERROR_ID : UINT;
END_VAR
VAR
  x : CW_REQUEST;
  prev : BOOL;
  refused : UINT;
  ms : UDINT;
  buf : ARRAY[0..1784] OF BYTE;
END_VAR
  ms := DWORD_TO_UDINT(TIME_TO_DWORD(TIMEOUT));
  IF ms > 65535 THEN
    ms := 65535;
  END_IF;
  IF EXECUTE AND NOT prev AND NOT x.BUSY THEN
    refused := 0;
    IF DESTINATION = 254 THEN
      refused := 3;
    END_IF;
  ELSIF NOT EXECUTE THEN
    refused := 0;
  END_IF;
  prev := EXECUTE;
  x(EXECUTE := EXECUTE AND refused = 0, OP := 14, NET := NETWORK, A0 := USINT_TO_WORD(DESTINATION),
    A1 := SEL(PREVIOUS_ONLY, WORD#0, WORD#1), A2 := UDINT_TO_WORD(ms), A3 := WORD#0, A4 := WORD#0, A5 := WORD#0, LENGTH := 0,
    FETCH_MAX := 0, LINK := LINK, DATA := buf);
  BUSY := x.BUSY;
  DONE := x.DONE;
  ERROR := x.ERROR OR refused <> 0;
  ERROR_ID := SEL(refused <> 0, x.ERROR_ID, refused);
END_FUNCTION_BLOCK

(* ---- J1939_DM_READ.st ---- *)
(*
 * J1939_DM_READ: the active trouble codes (DM1, PREVIOUS FALSE: the
 * bridge's latest DM1 from SOURCE, no bus traffic) or the previously active
 * ones (DM2, PREVIOUS TRUE: requested from SOURCE) of ECU SOURCE on J1939
 * network NETWORK: LAMPS and FLASH, COUNT codes in DTCS (up to 32), AGE of
 * the DM1. A rising edge of EXECUTE starts it; BUSY until the bridge has
 * an answer, then DONE or ERROR with ERROR_ID (docs/plc-library.md#j1939-blocks):
 * 1 the network is not running, 2 no such network, 3 invalid input,
 * 4 the network sends that PGN itself, 5 another DM2 read or clear for that
 * address is pending, 6 no answer within TIMEOUT, 7 the bus is off,
 * 8 cancelled, 9 no free job or receiver, 10 not a J1939 network, 11 the
 * network holds no address, 12 the destination answered NACK, 13 no DM1
 * from that source, 14 the transfer was aborted, 20 the bridge is not
 * reachable, 22 the config has no request mailbox.
 *)
(*
 * LINK is the generated `canworks.link` (ARRAY[0..1279] OF WORD); the block uses a request mailbox of the bridge (`mailboxes` in the config); instances share
 * them in the order they started (see
 * CW_LINK_SERVICE for the words).
 *)
FUNCTION_BLOCK J1939_DM_READ
VAR_INPUT
  EXECUTE : BOOL;
  NETWORK : USINT;
  SOURCE : USINT;
  PREVIOUS : BOOL;
  TIMEOUT : TIME;
END_VAR
VAR_IN_OUT
  DTCS : ARRAY[0..31] OF UDINT;
  LINK : ARRAY[0..1279] OF WORD;
END_VAR
VAR_OUTPUT
  BUSY : BOOL;
  DONE : BOOL;
  ERROR : BOOL;
  ERROR_ID : UINT;
  LAMPS : BYTE;
  FLASH : BYTE;
  COUNT : UINT;
  AGE : TIME;
END_VAR
VAR
  x : CW_REQUEST;
  prev : BOOL;
  refused : UINT;
  ms : UDINT;
  buf : ARRAY[0..1784] OF BYTE;
  was : BOOL;
  i : INT;
END_VAR
  ms := DWORD_TO_UDINT(TIME_TO_DWORD(TIMEOUT));
  IF ms > 65535 THEN
    ms := 65535;
  END_IF;
  IF EXECUTE AND NOT prev AND NOT x.BUSY THEN
    refused := 0;
    IF SOURCE > 253 THEN
      refused := 3;
    END_IF;
  ELSIF NOT EXECUTE THEN
    refused := 0;
  END_IF;
  prev := EXECUTE;
  x(EXECUTE := EXECUTE AND refused = 0, OP := 13, NET := NETWORK, A0 := USINT_TO_WORD(SOURCE),
    A1 := SEL(PREVIOUS, WORD#0, WORD#1), A2 := UDINT_TO_WORD(ms), A3 := WORD#0, A4 := WORD#0, A5 := WORD#0, LENGTH := 0,
    FETCH_MAX := 128, LINK := LINK, DATA := buf);
  BUSY := x.BUSY;
  DONE := x.DONE;
  ERROR := x.ERROR OR refused <> 0;
  ERROR_ID := SEL(refused <> 0, x.ERROR_ID, refused);
  IF x.DONE AND NOT was THEN
    LAMPS := WORD_TO_BYTE(SHR(x.R0, 8));
    FLASH := WORD_TO_BYTE(x.R0);
    COUNT := WORD_TO_UINT(x.R1);
    AGE := DWORD_TO_TIME(SHL(WORD_TO_DWORD(x.R2), 16) OR WORD_TO_DWORD(x.R3));
    FOR i := 0 TO 31 DO
      DTCS[i] := DWORD_TO_UDINT(SHL(BYTE_TO_DWORD(buf[4 * i]), 24) OR SHL(BYTE_TO_DWORD(buf[4 * i + 1]), 16) OR
                 SHL(BYTE_TO_DWORD(buf[4 * i + 2]), 8) OR BYTE_TO_DWORD(buf[4 * i + 3]));
    END_FOR;
  END_IF;
  was := x.DONE;
END_FUNCTION_BLOCK

(* ---- J1939_ECU_INFO.st ---- *)
(*
 * J1939_ECU_INFO: while ENABLE, the canworks ECU of J1939 network NETWORK
 * (one of the first 8) from the bridge's network info block, without a
 * request: VALID, STATE (0 claiming, 1 claimed, 2 cannot claim, 3 off),
 * ADDRESS, NAME, ECU_COUNT (ECUs seen on the bus). ERROR_ID
 * (docs/plc-library.md#j1939-blocks): 1 the network is not running, 2 no
 * such network, 10 not a J1939 network, 20 the bridge is not reachable,
 * 22 the config has no network info (or NETWORK is past the first 8).
 *)
(*
 * LINK is the generated `canworks.link` (ARRAY[0..1279] OF WORD); the block reads the bridge's network info block (see
 * CW_LINK_SERVICE for the words).
 *)
FUNCTION_BLOCK J1939_ECU_INFO
VAR_INPUT
  ENABLE : BOOL;
  NETWORK : USINT;
END_VAR
VAR_IN_OUT
  LINK : ARRAY[0..1279] OF WORD;
END_VAR
VAR_OUTPUT
  VALID : BOOL;
  STATE : USINT;
  ADDRESS : USINT;
  NAME : LWORD;
  ECU_COUNT : UINT;
  ERROR : BOOL;
  ERROR_ID : UINT;
END_VAR
VAR
  p : INT;
END_VAR
  ERROR_ID := 0;
  VALID := FALSE;
  IF NOT ENABLE THEN
    ERROR := FALSE;
    RETURN;
  END_IF;
  IF (LINK[21] AND WORD#16#0001) = WORD#0 THEN
    ERROR_ID := 20;
  ELSIF (LINK[89] AND WORD#16#0020) = WORD#0 OR NETWORK > 7 THEN
    ERROR_ID := 22;
  ELSE
    p := 960 + 18 * USINT_TO_INT(NETWORK);
    IF LINK[p + 17] = WORD#0 THEN
      ERROR_ID := 2;
    ELSIF SHR(LINK[p + 11], 8) = WORD#16#FF THEN
      ERROR_ID := WORD_TO_UINT(LINK[p + 11] AND WORD#16#00FF);
    END_IF;
  END_IF;
  ERROR := ERROR_ID <> 0;
  IF ERROR THEN
    STATE := 3;
    ADDRESS := 254;
    RETURN;
  END_IF;
  VALID := TRUE;
  STATE := WORD_TO_USINT(SHR(LINK[p + 11], 8));
  ADDRESS := WORD_TO_USINT(LINK[p + 11] AND WORD#16#00FF);
  NAME := SHL(WORD_TO_LWORD(LINK[p + 12]), 48) OR SHL(WORD_TO_LWORD(LINK[p + 13]), 32) OR
          SHL(WORD_TO_LWORD(LINK[p + 14]), 16) OR WORD_TO_LWORD(LINK[p + 15]);
  ECU_COUNT := WORD_TO_UINT(LINK[p + 16]);
END_FUNCTION_BLOCK

(* ---- J1939_FIND_ECU.st ---- *)
(*
 * J1939_FIND_ECU: while ENABLE, looks again and again on J1939 network
 * NETWORK for an ECU whose NAME matches NAME in the bits set in MASK
 * (FIND_ECU through a request mailbox; each look takes its turn): VALID
 * after the first answer, FOUND with its ADDRESS (254 when not found) and
 * FOUND_NAME, COUNT ECUs that match. ERROR_ID
 * (docs/plc-library.md#j1939-blocks): 1 the network is not running, 2 no
 * such network, 10 not a J1939 network, 20 the bridge is not reachable,
 * 22 the config has no request mailbox.
 *)
(*
 * LINK is the generated `canworks.link` (ARRAY[0..1279] OF WORD); the block uses a request mailbox of the bridge (`mailboxes` in the config); instances share
 * them in the order they started (see
 * CW_LINK_SERVICE for the words).
 *)
FUNCTION_BLOCK J1939_FIND_ECU
VAR_INPUT
  ENABLE : BOOL;
  NETWORK : USINT;
  NAME : LWORD;
  MASK : LWORD;
END_VAR
VAR_IN_OUT
  LINK : ARRAY[0..1279] OF WORD;
END_VAR
VAR_OUTPUT
  VALID : BOOL;
  FOUND : BOOL;
  ADDRESS : USINT;
  FOUND_NAME : LWORD;
  COUNT : UINT;
  ERROR : BOOL;
  ERROR_ID : UINT;
END_VAR
VAR
  x : CW_REQUEST;
  buf : ARRAY[0..1784] OF BYTE;
  run : BOOL;
  i : INT;
END_VAR
  IF NOT ENABLE THEN
    VALID := FALSE;
    FOUND := FALSE;
    ERROR := FALSE;
    ERROR_ID := 0;
    run := FALSE;
    x(EXECUTE := FALSE, LINK := LINK, DATA := buf);
    RETURN;
  END_IF;
  IF NOT x.BUSY THEN
    FOR i := 0 TO 7 DO
      buf[i] := LWORD_TO_BYTE(SHR(NAME, 56 - 8 * i));
      buf[8 + i] := LWORD_TO_BYTE(SHR(MASK, 56 - 8 * i));
    END_FOR;
  END_IF;
  (* One look per EXECUTE edge: the call after an answer drops it. *)
  run := NOT (x.DONE OR x.ERROR);
  x(EXECUTE := run, OP := 15, NET := NETWORK, A0 := WORD#0, A1 := WORD#0, A2 := WORD#0, A3 := WORD#0, A4 := WORD#0, A5 := WORD#0, LENGTH := 16,
    FETCH_MAX := 8, LINK := LINK, DATA := buf);
  IF x.DONE THEN
    VALID := TRUE;
    FOUND := x.R0 <> WORD#0;
    ADDRESS := SEL(FOUND, USINT#254, WORD_TO_USINT(x.R1));
    COUNT := WORD_TO_UINT(x.R2);
    FOUND_NAME := LWORD#0;
    FOR i := 0 TO 7 DO
      FOUND_NAME := SHL(FOUND_NAME, 8) OR BYTE_TO_LWORD(buf[i]);
    END_FOR;
    ERROR := FALSE;
    ERROR_ID := 0;
  ELSIF x.ERROR THEN
    VALID := FALSE;
    ERROR := TRUE;
    ERROR_ID := x.ERROR_ID;
  END_IF;
END_FUNCTION_BLOCK

(* ---- J1939_RECEIVE.st ---- *)
(*
 * J1939_RECEIVE: receives the messages of PGN (ALL_PGNS: every PGN) on J1939
 * network NETWORK, from SOURCE when FILTER_SOURCE, sent to the canworks ECU
 * or broadcast (ALL_DESTINATIONS: to any address), through a receiver of
 * the bridge with a queue of DEPTH messages (0: 4, at most 32). ENABLE
 * opens it; changed filter inputs open it again. Each call gives at most one
 * message, oldest first: RECEIVED with RX_PGN, RX_SOURCE, RX_DESTINATION,
 * RX_PRIORITY, RX_LENGTH bytes in RX_DATA and TIMESTAMP (UTC microseconds,
 * the receive time of the bridge's batch, which its messages share).
 * A message longer than 8 bytes is read whole (RX_FETCH through a request
 * mailbox) before RECEIVED. QUEUED messages still wait in the bridge, OVERFLOW
 * the queue was full, DROPPED messages lost. ERROR_ID
 * (docs/plc-library.md#j1939-blocks): 1 the network is not running, 2 no
 * such network, 3 invalid input, 8 the bridge closed the receiver (it opens
 * again), 9 no free receiver, 10 not a J1939 network, 20 the bridge is not
 * reachable, 22 the config has no receive or request mailbox. After 1, 8,
 * 9 and 20 it opens again by itself.
 *)
(*
 * LINK is the generated `canworks.link` (ARRAY[0..1279] OF WORD); the block uses the bridge's receive mailbox and a request mailbox (see
 * CW_LINK_SERVICE for the words).
 *)
FUNCTION_BLOCK J1939_RECEIVE
VAR_INPUT
  ENABLE : BOOL;
  NETWORK : USINT;
  PGN : UDINT;
  ALL_PGNS : BOOL;
  SOURCE : USINT;
  FILTER_SOURCE : BOOL;
  ALL_DESTINATIONS : BOOL;
  DEPTH : UINT;
END_VAR
VAR_IN_OUT
  RX_DATA : ARRAY[0..1784] OF BYTE;
  LINK : ARRAY[0..1279] OF WORD;
END_VAR
VAR_OUTPUT
  ACTIVE : BOOL;
  RECEIVED : BOOL;
  RX_PGN : UDINT;
  RX_SOURCE : USINT;
  RX_DESTINATION : USINT;
  RX_PRIORITY : USINT;
  RX_LENGTH : UINT;
  TIMESTAMP : ULINT;
  QUEUED : UINT;
  OVERFLOW : BOOL;
  DROPPED : UDINT;
  ERROR : BOOL;
  ERROR_ID : UINT;
END_VAR
VAR
  rx : CW_RX;
  fetch : CW_REQUEST;
  prev : BOOL;
  was_active : BOOL;
  fetching : BOOL;
  last_drop : WORD;
  src : USINT;
  flags : USINT;
  o_pgn : UDINT;
  o_source : USINT;
  o_flags : USINT;
  o_depth : UINT;
  changed : BOOL;
  rec : INT;
  i : INT;
  ferr : UINT;
END_VAR
  RECEIVED := FALSE;
  ferr := 0;
  IF ENABLE AND NOT prev THEN
    QUEUED := 0;
    OVERFLOW := FALSE;
    DROPPED := 0;
  END_IF;
  prev := ENABLE;
  src := SEL(FILTER_SOURCE, USINT#255, SOURCE);
  flags := SEL(ALL_PGNS, USINT#0, USINT#1) + SEL(ALL_DESTINATIONS, USINT#0, USINT#2);
  changed := rx.ACTIVE AND (PGN <> o_pgn OR src <> o_source OR flags <> o_flags OR DEPTH <> o_depth);
  IF NOT rx.ACTIVE THEN
    o_pgn := PGN;
    o_source := src;
    o_flags := flags;
    o_depth := DEPTH;
  END_IF;
  IF fetching THEN
    fetch(EXECUTE := TRUE, OP := 10, NET := NETWORK, A0 := INT_TO_WORD(rx.SLOT), A1 := WORD#0, A2 := WORD#0, A3 := WORD#0, A4 := WORD#0,
          A5 := WORD#0, LENGTH := 0, RLEN_AT := 0, FETCH_MAX := 1785, LINK := LINK, DATA := RX_DATA);
    IF fetch.DONE THEN
      fetching := FALSE;
      RECEIVED := TRUE;
      RX_LENGTH := fetch.GOT;
    ELSIF fetch.ERROR THEN
      fetching := FALSE;
      ferr := fetch.ERROR_ID;
    END_IF;
    IF NOT fetching THEN
      fetch(EXECUTE := FALSE, LINK := LINK, DATA := RX_DATA);
    END_IF;
  END_IF;
  rx(ENABLE := ENABLE, CHANGED := changed, NEXT := NOT fetching AND NOT RECEIVED, KIND := 2, NETWORK := NETWORK,
     FLAGS := flags, DEPTH := DEPTH, ID := PGN, MASK := USINT_TO_UDINT(src), RETRY := DWORD#16#00100302,
     LINK := LINK);
  IF rx.ACTIVE AND NOT was_active THEN
    last_drop := WORD#0;
  END_IF;
  was_active := rx.ACTIVE;
  IF rx.RECEIVED THEN
    rec := rx.REC;
    QUEUED := WORD_TO_UINT(LINK[rec + 1]);
    DROPPED := DROPPED + WORD_TO_UDINT(DINT_TO_WORD(WORD_TO_DINT(LINK[rec + 2]) - WORD_TO_DINT(last_drop)));
    last_drop := LINK[rec + 2];
    OVERFLOW := (LINK[rec] AND WORD#16#0004) <> WORD#0;
    TIMESTAMP := LWORD_TO_ULINT(SHL(WORD_TO_LWORD(LINK[741]), 48) OR SHL(WORD_TO_LWORD(LINK[742]), 32) OR
                 SHL(WORD_TO_LWORD(LINK[743]), 16) OR WORD_TO_LWORD(LINK[744]));
    RX_PGN := WORD_TO_UDINT(LINK[rec + 3]) * 65536 + WORD_TO_UDINT(LINK[rec + 4]);
    RX_SOURCE := WORD_TO_USINT(SHR(LINK[rec + 5], 8));
    RX_DESTINATION := WORD_TO_USINT(LINK[rec + 5] AND WORD#16#00FF);
    RX_PRIORITY := WORD_TO_USINT(LINK[rec + 6]);
    RX_LENGTH := WORD_TO_UINT(LINK[rec + 7]);
    IF (LINK[rec] AND WORD#16#0001) <> WORD#0 THEN
      (* Longer than 8 bytes: read it whole first. *)
      fetching := TRUE;
      fetch(EXECUTE := TRUE, OP := 10, NET := NETWORK, A0 := INT_TO_WORD(rx.SLOT), A1 := WORD#0, A2 := WORD#0, A3 := WORD#0,
            A4 := WORD#0, A5 := WORD#0, LENGTH := 0, RLEN_AT := 0, FETCH_MAX := 1785, LINK := LINK, DATA := RX_DATA);
    ELSE
      RECEIVED := TRUE;
      FOR i := 0 TO 3 DO
        RX_DATA[2 * i] := WORD_TO_BYTE(SHR(LINK[rec + 8 + i], 8));
        RX_DATA[2 * i + 1] := WORD_TO_BYTE(LINK[rec + 8 + i]);
      END_FOR;
    END_IF;
  END_IF;
  IF NOT rx.ACTIVE AND fetching THEN
    fetching := FALSE;
    fetch(EXECUTE := FALSE, LINK := LINK, DATA := RX_DATA);
  END_IF;
  ACTIVE := rx.ACTIVE;
  ERROR := rx.ERROR OR ferr <> 0;
  ERROR_ID := SEL(ferr <> 0, rx.ERROR_ID, ferr);
END_FUNCTION_BLOCK

(* ---- J1939_REQUEST.st ---- *)
(*
 * J1939_REQUEST: requests PGN from DESTINATION (255: every ECU, the first
 * answer counts) on J1939 network NETWORK and returns the answer: SOURCE,
 * LENGTH bytes in DATA (up to 1785), ACK_CODE of an acknowledgement. A rising edge of EXECUTE starts it; BUSY until the bridge has
 * an answer, then DONE or ERROR with ERROR_ID (docs/plc-library.md#j1939-blocks):
 * 1 the network is not running, 2 no such network, 3 invalid input,
 * 4 the network sends that PGN itself, 5 another DM2 read or clear for that
 * address is pending, 6 no answer within TIMEOUT, 7 the bus is off,
 * 8 cancelled, 9 no free job or receiver, 10 not a J1939 network, 11 the
 * network holds no address, 12 the destination answered NACK, 13 no DM1
 * from that source, 14 the transfer was aborted, 20 the bridge is not
 * reachable, 22 the config has no request mailbox.
 *)
(*
 * LINK is the generated `canworks.link` (ARRAY[0..1279] OF WORD); the block uses a request mailbox of the bridge (`mailboxes` in the config); instances share
 * them in the order they started (see
 * CW_LINK_SERVICE for the words).
 *)
FUNCTION_BLOCK J1939_REQUEST
VAR_INPUT
  EXECUTE : BOOL;
  NETWORK : USINT;
  PGN : UDINT;
  DESTINATION : USINT;
  TIMEOUT : TIME;
END_VAR
VAR_IN_OUT
  DATA : ARRAY[0..1784] OF BYTE;
  LINK : ARRAY[0..1279] OF WORD;
END_VAR
VAR_OUTPUT
  BUSY : BOOL;
  DONE : BOOL;
  ERROR : BOOL;
  ERROR_ID : UINT;
  SOURCE : USINT;
  LENGTH : UINT;
  ACK_CODE : USINT;
END_VAR
VAR
  x : CW_REQUEST;
  prev : BOOL;
  refused : UINT;
  ms : UDINT;
  was : BOOL;
END_VAR
  ms := DWORD_TO_UDINT(TIME_TO_DWORD(TIMEOUT));
  IF ms > 65535 THEN
    ms := 65535;
  END_IF;
  IF EXECUTE AND NOT prev AND NOT x.BUSY THEN
    refused := 0;
    ACK_CODE := 0;
  ELSIF NOT EXECUTE THEN
    refused := 0;
  END_IF;
  prev := EXECUTE;
  x(EXECUTE := EXECUTE AND refused = 0, OP := 12, NET := NETWORK, A0 := DWORD_TO_WORD(SHR(UDINT_TO_DWORD(PGN), 16)),
    A1 := UDINT_TO_WORD(PGN), A2 := USINT_TO_WORD(DESTINATION), A3 := UDINT_TO_WORD(ms), A4 := WORD#0, A5 := WORD#0,
    LENGTH := 0, RLEN_AT := 1, FETCH_MAX := 1785, LINK := LINK, DATA := DATA);
  BUSY := x.BUSY;
  DONE := x.DONE;
  ERROR := x.ERROR OR refused <> 0;
  ERROR_ID := SEL(refused <> 0, x.ERROR_ID, refused);
  IF (x.DONE OR x.ERROR) AND NOT was THEN
    ACK_CODE := WORD_TO_USINT(x.R2);
    IF x.DONE THEN
      SOURCE := WORD_TO_USINT(x.R0);
      LENGTH := WORD_TO_UINT(x.R1);
    END_IF;
  END_IF;
  was := x.DONE OR x.ERROR;
END_FUNCTION_BLOCK

(* ---- J1939_SEND.st ---- *)
(*
 * J1939_SEND: sends LENGTH bytes of DATA (0..1785; more than 8 by the
 * transport protocol, BAM to 255) as PGN to DESTINATION with PRIORITY (0: 6)
 * on J1939 network NETWORK. A rising edge of EXECUTE starts it; BUSY until the bridge has
 * an answer, then DONE or ERROR with ERROR_ID (docs/plc-library.md#j1939-blocks):
 * 1 the network is not running, 2 no such network, 3 invalid input,
 * 4 the network sends that PGN itself, 5 another DM2 read or clear for that
 * address is pending, 6 no answer within TIMEOUT, 7 the bus is off,
 * 8 cancelled, 9 no free job or receiver, 10 not a J1939 network, 11 the
 * network holds no address, 12 the destination answered NACK, 13 no DM1
 * from that source, 14 the transfer was aborted, 20 the bridge is not
 * reachable, 22 the config has no request mailbox.
 *)
(*
 * LINK is the generated `canworks.link` (ARRAY[0..1279] OF WORD); the block uses a request mailbox of the bridge (`mailboxes` in the config); instances share
 * them in the order they started (see
 * CW_LINK_SERVICE for the words).
 *)
FUNCTION_BLOCK J1939_SEND
VAR_INPUT
  EXECUTE : BOOL;
  NETWORK : USINT;
  PGN : UDINT;
  DESTINATION : USINT;
  PRIORITY : USINT;
  LENGTH : UINT;
  TIMEOUT : TIME;
END_VAR
VAR_IN_OUT
  DATA : ARRAY[0..1784] OF BYTE;
  LINK : ARRAY[0..1279] OF WORD;
END_VAR
VAR_OUTPUT
  BUSY : BOOL;
  DONE : BOOL;
  ERROR : BOOL;
  ERROR_ID : UINT;
END_VAR
VAR
  x : CW_REQUEST;
  prev : BOOL;
  refused : UINT;
  ms : UDINT;
  prio : USINT;
END_VAR
  ms := DWORD_TO_UDINT(TIME_TO_DWORD(TIMEOUT));
  IF ms > 65535 THEN
    ms := 65535;
  END_IF;
  IF EXECUTE AND NOT prev AND NOT x.BUSY THEN
    refused := 0;
    IF LENGTH > 1785 OR PRIORITY > 7 THEN
      refused := 3;
    END_IF;
  ELSIF NOT EXECUTE THEN
    refused := 0;
  END_IF;
  prev := EXECUTE;
  prio := PRIORITY;
  IF prio = 0 THEN
    prio := 6;
  END_IF;
  x(EXECUTE := EXECUTE AND refused = 0, OP := 11, NET := NETWORK, A0 := DWORD_TO_WORD(SHR(UDINT_TO_DWORD(PGN), 16)),
    A1 := UDINT_TO_WORD(PGN), A2 := SHL(USINT_TO_WORD(DESTINATION), 8) OR USINT_TO_WORD(prio),
    A3 := UINT_TO_WORD(LENGTH), A4 := UDINT_TO_WORD(ms), A5 := WORD#0, LENGTH := LENGTH, FETCH_MAX := 0, LINK := LINK,
    DATA := DATA);
  BUSY := x.BUSY;
  DONE := x.DONE;
  ERROR := x.ERROR OR refused <> 0;
  ERROR_ID := SEL(refused <> 0, x.ERROR_ID, refused);
END_FUNCTION_BLOCK
